(* IEC 61131-3 sources: daoli-st-library/DL_Device (part 28) *)

(* ---- FB_DL_PneumaticCylinder.st ---- *)
(*==============================================================================
 * 组件名称 (Component)  : FB_DL_PneumaticCylinder
 * 所属子库 (Sublibrary) : DL_Device
 * 当前版本 (Version)    : 1.0.1
 * 兼容性   (Platform)   : CODESYS 3.5 / TwinCAT 3 / 汇川 InoProShop / Machine Expert
 *                         仅依赖 Standard.library（TON / R_TRIG）与本库 DL_Base
 *                         的 FB_DL_SignalDebounce，零厂商方言
 * 分类     (Category)   : 设备执行器功能块（Function Block，实现 I_DL_Cylinder）
 * 功能简述 (Function)   : 标准双电控（双线圈）气缸控制功能块。含磁开信号双通道
 *                         消抖、伸出/缩回超时自检、双传感器位置冲突锁存、
 *                         双线圈互斥出口断言、联锁失电保位、行程计数；
 *                         状态机采用 ENUM + CASE + ELSE 兜底。
 * 接口实现 (Implements) : I_DL_Cylinder（属性 eState/bExtended/bRetracted/
 *                         bFault/uErrorId，方法 CmdExtend/CmdRetract/
 *                         CmdStop/CmdReset，全部在本文件尾部落地）
 * 开源溯源 (Origin)     : 来源标签 lbp-device（RAW_NOTES_R5 S-4：工业气动气缸
 *                         FB 设计指南 / 双电控 5/2 阀 + 磁性开关 + 行程计数
 *                         接线语义 / 双线圈禁止同时得电互锁惯例，公开教学
 *                         文章，仅借鉴通用工程语义；状态机、故障码、互斥
 *                         断言按本库红线独立设计，clean-room 未复制源码）。
 * 红线自检 (Redline)    : R1 零全局变量表/外部变量引用 ✓｜R2 零物理 IO 地址 ✓
 *                         R3 纯 IEC 61131-3 ✓｜R4 防越界/互斥断言 ✓
 *                         R5 全变量中英双语同行注释 ✓｜R6 ENUM+CASE+ELSE ✓
 *                         R7 六个定时器/边缘实例主体最前部无条件刷新 ✓
 * 公约遵循 (Convention) : 0.1 本块为纯事件型状态机，无积分/滤波类首扫初始化
 *                         逻辑（消抖由 FB_DL_SignalDebounce 内部自理），
 *                         首扫跟踪范式不适用，无内部初始化标志。
 *                         0.7 故障码段位 16#0003_xxxx：0003_0201 非法状态/
 *                         0003_0202 伸出超时/0003_0203 缩回超时/0003_0204
 *                         双传感器冲突，全部【故障级】R15 锁存仅复位可清；
 *                         本块无信息级码，bFault 派生式天然排除信息级（0.2）。
 * 修订历史 (Revision)   :
 *   2026-11-15  v1.0.0  首版入库（R5 轮 · DL_Device 开库）
 *   2026-11-15  v1.0.1  R11 修复：变量名勘误，段 2 行程计数赋值目标
 *                       _uCycleCount → uCycleCount（原写下划线前缀但未在
 *                       VAR 区声明，且同名输出 uCycleCount 全文零写入，
 *                       判定为前缀笔误而非缺声明；三平台编译阻断已消除）。
 *                       R11 fix: name erratum, _uCycleCount -> uCycleCount
 *============================================================================*)
FUNCTION_BLOCK FB_DL_PneumaticCylinder IMPLEMENTS I_DL_Cylinder
VAR_INPUT
    bCmdExtend    : BOOL;         // 伸出指令（Extend command），上升沿生效 / Extend command, rising edge effective
    bCmdRetract   : BOOL;         // 缩回指令（Retract command），上升沿生效 / Retract command, rising edge effective
    bSnsExtended  : BOOL;         // 伸出到位磁性开关（Extended reed switch），TRUE=到位 / Extended reed switch, TRUE = in position
    bSnsRetracted : BOOL;         // 缩回到位磁性开关（Retracted reed switch），TRUE=到位 / Retracted reed switch, TRUE = in position
    bInterlock    : BOOL;         // 允许动作联锁（Motion interlock），TRUE=允许动作，默认 FALSE 双线圈保持断开 / Motion interlock, TRUE = motion allowed, default FALSE holds coils off
    tTimeoutExt   : TIME := T#2S; // 伸出到位超时（Extend timeout），T#0S=禁用自检 / Extend timeout, T#0S disables the check
    tTimeoutRet   : TIME := T#2S; // 缩回到位超时（Retract timeout），T#0S=禁用自检 / Retract timeout, T#0S disables the check
    tDebounce     : TIME := T#20MS; // 磁开防抖窗口（Sensor debounce），T#0S=直通 / Sensor debounce window, T#0S = pass-through
    bReset        : BOOL;         // 故障复位（Fault reset），上升沿生效 / Fault reset, rising edge effective
END_VAR

VAR_OUTPUT
    bSolenoidExt  : BOOL;         // 伸出线圈输出（Extend solenoid coil），TRUE=得电 / Extend solenoid coil, TRUE = energized
    bSolenoidRet  : BOOL;         // 缩回线圈输出（Retract solenoid coil），TRUE=得电 / Retract solenoid coil, TRUE = energized
    eState        : E_DL_CylinderState; // 当前状态机状态（Current state），映射接口同名属性 / Current state, mirrors interface property
    bExtended     : BOOL;         // 伸出到位磁开反馈（Extended reed feedback），消抖后 / Extended reed feedback, debounced
    bRetracted    : BOOL;         // 缩回到位磁开反馈（Retracted reed feedback），消抖后 / Retracted reed feedback, debounced
    bMoving       : BOOL;         // 运动中指示（Moving indicator），TRUE=伸出或缩回动作中 / Moving indicator, TRUE while extending or retracting
    bFault        : BOOL;         // 故障锁存中（Fault latched），TRUE=需复位 / Fault latched, TRUE requires reset
    uErrorId      : UDINT;        // 末次故障码（Last error code），0=无故障，段位 16#0003_xxxx / Last error code, 0 = none, family 16#0003_xxxx
    uCycleCount   : UDINT;        // 行程计数（Stroke count），缩回到位上升沿 +1 / Stroke count, incremented on retracted-position rising edge
END_VAR

VAR
    _eState       : E_DL_CylinderState := E_DL_CylinderState.eIdle; // 内部状态机步序（Internal state step），外部经属性只读 / Internal state, read-only via property
    _bFaultLatch  : BOOL;         // 故障锁存标志（Fault latch flag），仅复位清除 / Fault latch flag, cleared only by reset
    _uErrorIdInt  : UDINT;        // 内部故障码寄存（Internal error register），随锁存写入 / Internal error register written on latch
    _bPendExtend  : BOOL;         // 方法伸出请求锁存（Method extend request），由 CmdExtend 置位 / Method extend request set by CmdExtend
    _bPendRetract : BOOL;         // 方法缩回请求锁存（Method retract request），由 CmdRetract 置位 / Method retract request set by CmdRetract
    _bPendStop    : BOOL;         // 方法停止请求锁存（Method stop request），由 CmdStop 置位 / Method stop request set by CmdStop
    _bPendReset   : BOOL;         // 方法复位请求锁存（Method reset request），由 CmdReset 置位 / Method reset request set by CmdReset
    _bExtFilt     : BOOL;         // 消抖后伸出磁开（Debounced extended reed）/ Debounced extended reed signal
    _bRetFilt     : BOOL;         // 消抖后缩回磁开（Debounced retracted reed）/ Debounced retracted reed signal
    _bExtToEn     : BOOL;         // 伸出超时自检使能（Extend timeout check enable），超时参数大于零时有效 / Extend timeout enable, active when timeout parameter above zero
    _bRetToEn     : BOOL;         // 缩回超时自检使能（Retract timeout check enable），超时参数大于零时有效 / Retract timeout enable, active when timeout parameter above zero
    _fbDebExt     : FB_DL_SignalDebounce; // 伸出磁开消抖实例（Extended reed debounce），通道一 / Extended reed debounce instance, channel 1
    _fbDebRet     : FB_DL_SignalDebounce; // 缩回磁开消抖实例（Retracted reed debounce），通道二 / Retracted reed debounce instance, channel 2
    _fbTrigExt    : R_TRIG;       // 引脚伸出指令上升沿（Pin extend command edge）/ Pin extend command rising edge
    _fbTrigRet    : R_TRIG;       // 引脚缩回指令上升沿（Pin retract command edge）/ Pin retract command rising edge
    _fbTrigReset  : R_TRIG;       // 引脚复位上升沿（Pin reset edge）/ Pin reset rising edge
    _fbTrigStroke : R_TRIG;       // 缩回到位计数上升沿（Stroke count edge）/ Stroke count rising edge on retracted feedback
    _fbTonExtTo   : TON;          // 伸出到位超时定时器（Extend timeout timer）/ Extend timeout timer instance
    _fbTonRetTo   : TON;          // 缩回到位超时定时器（Retract timeout timer）/ Retract timeout timer instance
END_VAR

METHOD CmdExtend : BOOL
VAR_INPUT
END_VAR
IF _bFaultLatch OR (_eState = E_DL_CylinderState.eFault) THEN
    CmdExtend     := FALSE;   // 故障态拒绝（Rejected in fault state）
    _bPendRetract := FALSE;   // 清反向残留请求（Clear stale reverse request）
ELSE
    _bPendExtend  := TRUE;    // 登记伸出请求（Register extend request）
    _bPendRetract := FALSE;   // 互斥注销反向请求（Cancel opposite request）
    CmdExtend     := TRUE;    // 受理成功（Accepted）
END_IF

(*------------------------------------------------------------------------------
 * 方法: CmdRetract —— 缩回指令（单发）。故障锁存态一律拒绝并返回 FALSE。
 *      Method CmdRetract - retract command (one-shot), rejected with FALSE in fault state.
 *------------------------------------------------------------------------------*)
    END_METHOD

METHOD CmdRetract : BOOL
VAR_INPUT
END_VAR
IF _bFaultLatch OR (_eState = E_DL_CylinderState.eFault) THEN
    CmdRetract   := FALSE;    // 故障态拒绝（Rejected in fault state）
    _bPendExtend := FALSE;    // 清反向残留请求（Clear stale reverse request）
ELSE
    _bPendRetract := TRUE;    // 登记缩回请求（Register retract request）
    _bPendExtend  := FALSE;   // 互斥注销反向请求（Cancel opposite request）
    CmdRetract    := TRUE;    // 受理成功（Accepted）
END_IF

(*------------------------------------------------------------------------------
 * 方法: CmdStop —— 双线圈全断、保持当前位置。故障锁存态拒绝返回 FALSE。
 *      Method CmdStop - both coils off and hold position, rejected with FALSE in fault state.
 *------------------------------------------------------------------------------*)
    END_METHOD

METHOD CmdStop : BOOL
VAR_INPUT
END_VAR
IF _bFaultLatch OR (_eState = E_DL_CylinderState.eFault) THEN
    CmdStop := FALSE;         // 故障态拒绝（Rejected in fault state）
ELSE
    _bPendExtend  := FALSE;   // 注销全部动作请求（Cancel all motion requests）
    _bPendRetract := FALSE;
    _bPendStop    := TRUE;    // 登记停止请求，主体状态机消化（Register stop request, consumed by body）
    CmdStop       := TRUE;    // 受理成功（Accepted）
END_IF

(*------------------------------------------------------------------------------
 * 方法: CmdReset —— 复位故障，返回是否可复位（存在锁存故障时为 TRUE）。
 *      Method CmdReset - reset fault, returns TRUE only when a latch exists.
 *------------------------------------------------------------------------------*)
    END_METHOD

METHOD CmdReset : BOOL
VAR_INPUT
END_VAR
IF _bFaultLatch OR (_eState = E_DL_CylinderState.eFault) THEN
    _bPendReset := TRUE;      // 登记复位请求，主体状态机消化（Register reset request, consumed by body）
    CmdReset    := TRUE;      // 可复位（Resettable）
ELSE
    CmdReset    := FALSE;     // 无故障可复位（Nothing to reset）
END_IF

(*------------------------------------------------------------------------------
 * 属性: eState（GET）—— 当前状态机状态只读视图。
 *      Property eState (GET) - read-only view of the current state machine state.
 *------------------------------------------------------------------------------*)
    END_METHOD

// ============================================================================
// 段 1｜定时器与边缘检测实例无条件周期刷新（R7：严禁置于 IF/CASE 分支内）
//      Unconditional per-cycle refresh of all timer and edge instances (R7)
// ============================================================================
_fbDebExt(bRawInput := bSnsExtended, tRiseDelay := tDebounce, tFallDelay := tDebounce, bEnable := TRUE, bReset := FALSE);
_fbDebRet(bRawInput := bSnsRetracted, tRiseDelay := tDebounce, tFallDelay := tDebounce, bEnable := TRUE, bReset := FALSE);
_fbTrigExt(CLK := bCmdExtend);
_fbTrigRet(CLK := bCmdRetract);
_fbTrigReset(CLK := bReset);
_bExtFilt := _fbDebExt.bStable;   // 通道一消抖输出（Channel 1 debounced output）
_bRetFilt := _fbDebRet.bStable;   // 通道二消抖输出（Channel 2 debounced output）
_fbTrigStroke(CLK := _bRetFilt);

_bExtToEn := (tTimeoutExt > T#0S); // 超时参数为零 = 自检禁用（Zero timeout = check disabled）
_bRetToEn := (tTimeoutRet > T#0S); // 超时参数为零 = 自检禁用（Zero timeout = check disabled）
_fbTonExtTo(IN := (_eState = E_DL_CylinderState.eExtending) AND _bExtToEn, PT := tTimeoutExt);
_fbTonRetTo(IN := (_eState = E_DL_CylinderState.eRetracting) AND _bRetToEn, PT := tTimeoutRet);

// ============================================================================
// 段 2｜行程计数：缩回到位上升沿 +1（R15 范畴外，非故障量，不锁存）
//      Stroke counting: one increment per retracted-position rising edge
// ============================================================================
IF _fbTrigStroke.Q THEN
    uCycleCount := uCycleCount + 1; // 完整行程 +1（One completed stroke added）
END_IF

// ============================================================================
// 段 3｜位置冲突全局监视：双磁开同时动作物理不可能，立即锁存（优先级最高）
//      Global position-conflict monitor: both reed switches ON is physically
//      impossible, latch immediately (highest priority over the state machine)
// ============================================================================
IF _bExtFilt AND _bRetFilt THEN
    _bFaultLatch := TRUE;                          // 故障锁存（Fault latched）
    _uErrorIdInt := 16#0003_0204;                  // 0003_0204 双传感器同时动作【故障级】/ Both sensors active, fault level
    _eState      := E_DL_CylinderState.eFault;     // 强制进入故障态（Force fault state）
END_IF

// ============================================================================
// 段 4｜核心状态机（ENUM + CASE，含 ELSE 非法状态兜底）
//      Core state machine (ENUM + CASE with ELSE illegal-state fallback)
// ============================================================================
CASE _eState OF

    E_DL_CylinderState.eIdle: // 空闲稳态：双线圈全断，按传感器同步实际位置
        IF _bExtFilt AND (NOT _bRetFilt) THEN
            _eState := E_DL_CylinderState.eExtended;  // 首态同步：实际已伸出（Sync: physically extended）
        ELSIF _bRetFilt AND (NOT _bExtFilt) THEN
            _eState := E_DL_CylinderState.eRetracted; // 首态同步：实际已缩回（Sync: physically retracted）
        ELSIF (_bPendExtend OR _fbTrigExt.Q) AND bInterlock THEN
            _bPendExtend  := FALSE;                    // 消费伸出请求（Consume extend request）
            _eState       := E_DL_CylinderState.eExtending;
        ELSIF (_bPendRetract OR _fbTrigRet.Q) AND bInterlock THEN
            _bPendRetract := FALSE;                    // 消费缩回请求（Consume retract request）
            _eState       := E_DL_CylinderState.eRetracting;
        ELSIF _bPendStop THEN
            _bPendStop := FALSE;                       // 空闲态停止请求直接消化（Stop request absorbed in idle）
        END_IF

    E_DL_CylinderState.eExtending: // 伸出动作中：伸出线圈得电
        IF _bExtFilt AND (NOT _bRetFilt) THEN
            _eState := E_DL_CylinderState.eExtended;   // 到位确认（Reached extended position）
        ELSIF _fbTonExtTo.Q THEN
            _bFaultLatch := TRUE;                      // 超时故障锁存（Timeout fault latch）
            _uErrorIdInt := 16#0003_0202;              // 0003_0202 伸出到位超时【故障级】/ Extend timeout, fault level
            _eState      := E_DL_CylinderState.eFault;
        ELSIF NOT bInterlock THEN
            _eState := E_DL_CylinderState.eIdle;       // 联锁中途撤除：双线圈断、保位、不判故障（Interlock dropped mid-stroke: coils off, hold position, no fault）
        ELSIF _bPendStop THEN
            _bPendStop := FALSE;                       // 停止指令：双线圈全断保位（Stop command: both coils off, hold position）
            _eState    := E_DL_CylinderState.eIdle;
        ELSIF (_bPendRetract OR _fbTrigRet.Q) AND bInterlock THEN
            _bPendRetract := FALSE;                    // 行程中途反向（Mid-stroke reversal to retract）
            _eState       := E_DL_CylinderState.eRetracting;
        END_IF

    E_DL_CylinderState.eExtended: // 已伸出到位稳态
        IF _bPendStop THEN
            _bPendStop := FALSE;                       // 停止请求消化（Stop request absorbed）
            _eState    := E_DL_CylinderState.eIdle;
        ELSIF (_bPendRetract OR _fbTrigRet.Q) AND bInterlock THEN
            _bPendRetract := FALSE;                    // 受理缩回（Accept retract command）
            _eState       := E_DL_CylinderState.eRetracting;
        END_IF

    E_DL_CylinderState.eRetracting: // 缩回动作中：缩回线圈得电
        IF _bRetFilt AND (NOT _bExtFilt) THEN
            _eState := E_DL_CylinderState.eRetracted;  // 到位确认（Reached retracted position）
        ELSIF _fbTonRetTo.Q THEN
            _bFaultLatch := TRUE;                      // 超时故障锁存（Timeout fault latch）
            _uErrorIdInt := 16#0003_0203;              // 0003_0203 缩回到位超时【故障级】/ Retract timeout, fault level
            _eState      := E_DL_CylinderState.eFault;
        ELSIF NOT bInterlock THEN
            _eState := E_DL_CylinderState.eIdle;       // 联锁中途撤除：双线圈断、保位、不判故障（Interlock dropped mid-stroke: coils off, hold position, no fault）
        ELSIF _bPendStop THEN
            _bPendStop := FALSE;                       // 停止指令：双线圈全断保位（Stop command: both coils off, hold position）
            _eState    := E_DL_CylinderState.eIdle;
        ELSIF (_bPendExtend OR _fbTrigExt.Q) AND bInterlock THEN
            _bPendExtend := FALSE;                     // 行程中途反向（Mid-stroke reversal to extend）
            _eState      := E_DL_CylinderState.eExtending;
        END_IF

    E_DL_CylinderState.eRetracted: // 已缩回到位稳态
        IF _bPendStop THEN
            _bPendStop := FALSE;                       // 停止请求消化（Stop request absorbed）
            _eState    := E_DL_CylinderState.eIdle;
        ELSIF (_bPendExtend OR _fbTrigExt.Q) AND bInterlock THEN
            _bPendExtend := FALSE;                     // 受理伸出（Accept extend command）
            _eState      := E_DL_CylinderState.eExtending;
        END_IF

    E_DL_CylinderState.eFault: // 故障锁存态：清空全部请求，仅复位可退出
        _bPendExtend  := FALSE;                        // 清方法请求（Clear method requests）
        _bPendRetract := FALSE;
        _bPendStop    := FALSE;
        IF _bPendReset OR _fbTrigReset.Q THEN
            _bPendReset  := FALSE;                     // 消费复位请求（Consume reset request）
            _bFaultLatch := FALSE;                     // 解除锁存（Release latch）
            _uErrorIdInt := 0;                         // 故障码清零（Error code cleared）
            _eState      := E_DL_CylinderState.eIdle;  // 回空闲态重新同步（Back to idle for re-sync）
        END_IF

    ELSE // 非法状态兜底：任何越界枚举值强制锁存故障（Illegal state fallback）
        _bFaultLatch := TRUE;                          // 故障锁存（Fault latched）
        _uErrorIdInt := 16#0003_0201;                  // 0003_0201 非法状态【故障级】/ Illegal state, fault level
        _eState      := E_DL_CylinderState.eFault;
END_CASE

// ============================================================================
// 段 5｜线圈输出推导 + 双线圈互斥出口断言（硬约束：两输出恒不可同真）
//      Coil output derivation + dual-coil exclusivity assertion at exit
// ============================================================================
bSolenoidExt := (_eState = E_DL_CylinderState.eExtending);   // 仅动作态单端置位（Energize only during motion）
bSolenoidRet := (_eState = E_DL_CylinderState.eRetracting);
IF bSolenoidExt AND bSolenoidRet THEN
    bSolenoidExt := FALSE;                                   // 断言对调：异常同真时双断保安全（Assertion fallback: cut both on impossible condition）
    bSolenoidRet := FALSE;
END_IF

// ============================================================================
// 段 6｜状态引脚映射（bFault 为显式派生式，排除信息级码——本块无信息级码）
//      Status pin mapping (bFault explicit derived form, info codes excluded)
// ============================================================================
eState     := _eState;                                       // 状态映射（State mapping）
bExtended  := _bExtFilt;                                     // 伸出反馈映射（Extended feedback mapping）
bRetracted := _bRetFilt;                                     // 缩回反馈映射（Retracted feedback mapping）
bMoving    := (_eState = E_DL_CylinderState.eExtending) OR (_eState = E_DL_CylinderState.eRetracting); // 运动中派生（Moving derived）
bFault     := _bFaultLatch OR (_eState = E_DL_CylinderState.eFault); // 故障派生（Fault derived）
uErrorId   := _uErrorIdInt;                                  // 故障码映射（Error code mapping）

(*------------------------------------------------------------------------------
 * 方法: CmdExtend —— 伸出指令（单发）。故障锁存态一律拒绝并返回 FALSE。
 *      Method CmdExtend - extend command (one-shot), rejected with FALSE in fault state.
 *------------------------------------------------------------------------------*)

PROPERTY eState : E_DL_CylinderState
eState := _eState;            // 返回内部状态（Return internal state）

(*------------------------------------------------------------------------------
 * 属性: bExtended（GET）—— 伸出到位磁开反馈（消抖后）。
 *      Property bExtended (GET) - debounced extended reed feedback.
 *------------------------------------------------------------------------------*)
PROPERTY bExtended : BOOL
bExtended := _bExtFilt;       // 返回通道一消抖输出（Return channel 1 debounced output）

(*------------------------------------------------------------------------------
 * 属性: bRetracted（GET）—— 缩回到位磁开反馈（消抖后）。
 *      Property bRetracted (GET) - debounced retracted reed feedback.
 *------------------------------------------------------------------------------*)
PROPERTY bRetracted : BOOL
bRetracted := _bRetFilt;      // 返回通道二消抖输出（Return channel 2 debounced output）

(*------------------------------------------------------------------------------
 * 属性: bFault（GET）—— 故障锁存指示（信息级码不置本位，0.2 公约）。
 *      Property bFault (GET) - fault latch indicator, info-level codes excluded.
 *------------------------------------------------------------------------------*)
PROPERTY bFault : BOOL
bFault := _bFaultLatch OR (_eState = E_DL_CylinderState.eFault); // 显式排除信息级派生式（Explicit derived form excluding info codes）

(*------------------------------------------------------------------------------
 * 属性: uErrorId（GET）—— 末次故障码（0=无故障）。
 *      Property uErrorId (GET) - last error code (0 = none).
 *------------------------------------------------------------------------------*)
PROPERTY uErrorId : UDINT
uErrorId := _uErrorIdInt;     // 返回内部故障码寄存（Return internal error register）
END_FUNCTION_BLOCK

(* ---- FB_DL_PouchSwellingGauge.st ---- *)
(*
  FB_DL_PouchSwellingGauge  —  软包电芯鼓胀厚度巡检分级 / Pouch cell swelling thickness gauge and grading
  分类 Category : DL_Device
  码位 Code     : 16#03_2_15
  段位说明      : 03_2 段低半字节 00~0F 已满（05 为历史空穴留存），进位 15 段续号（R192）
  版本 Version  : 1.0.0
  来源 Source   : t2-1-lgf-measurement — IEC 61131-3 标准语义的道莅防御性实现
  溯源 Origin   : clean-room 实现，Welford 在线方差递推公开算法语义，未复制任何源码行
                  （统计语义对齐 FB_DL_SignalStatistics；分级语义对齐 FC_DL_LimitClassify，均不实例化）
  功能 Function : 1) 厚度归一（fThicknessMm − fZeroOffsetMm）后按批 Welford 递推均值/标准差（防大数累加误差）；
                  2) 单件双口径分级：绝对限 fAbsLimitMm 与 Z 分数 |x − mean|/σ > fZScoreLimit，越限立置 abItemNg[k]；
                  3) 批内一致性评价：σ > fBatchSigmaLimitMm 判 bBatchAbnormal（判据取「批内异常」而非单件越限）；
                  4) 批尾自动清零（计数/均值/NG 位全清，下批重来）。
  边界 Boundary : ① fAbsLimitMm <= 0 或 nBatchSize < 2（无法算 σ）判组态错；
                  ② nBatchSize > 数组上界按 MIN 钳制并置信息码（禁 TRUNC(x)+1 型写法，R28-2）；
                  ③ 批内 σ < 1E-6 mm 时 Z 分数不计算、只走绝对限（防除零）；
                  ④ fThicknessMm 非有限（NaN 用 x<>x 自反）判信号无效置码且不纳入统计（不污染均值）；
                  ⑤ 单件越限立刻置 abItemNg[k] 且本件锁存至批尾（解除式 = 批尾清零，可由 nBatchSize 满足）；
                  ⑥ 无状态机：统计件无 ENUM/CASE，判据均为每拍重算或批内锁存（批尾清零承载解除）。
  依赖 Depends  : 仅 Standard.library（ABS/SQRT/MIN）；语义对齐 FB_DL_SignalStatistics / FC_DL_LimitClassify（已注册）
  码表 Error codes（本件格 03_2_15，子码步进 +0x100）:
    16#0003_0115 信息级：批尾清零（批次评价已给出，不置故障）
    16#0003_0215 故障级：组态非法（绝对限 <= 0 / 批容量 < 2）
    16#0003_0315 信息级：批容量超数组上界，已按 MIN 钳制
    16#0003_0415 信息级：测量值非有限（NaN/Inf），本件不纳入统计
    16#0003_0515 信息级：批内 σ 近零，Z 分数不计算只走绝对限
    16#0003_0615 故障级：批内异常（σ 越限，批内一致性判废）

  修订历史 Revision :
    2026-11-18  v1.0.0  R38 首版
*)

FUNCTION_BLOCK FB_DL_PouchSwellingGauge
VAR_INPUT
    fThicknessMm       : REAL := 0.0;      // 测厚原始值 [mm] / Raw thickness measurement
    fZeroOffsetMm      : REAL := 0.0;      // 零点偏移 [mm] / Zero offset
    fAbsLimitMm        : REAL := 5.0;      // 绝对上限 [mm]，域 > 0 / Absolute thickness ceiling
    nBatchSize         : INT   := 32;      // 批内样本数上限 [件]，域 >= 2 / Batch size ceiling
    fBatchSigmaLimitMm : REAL := 0.05;     // 批内离散度上限 [mm]，域 > 0 / Batch sigma limit
    fZScoreLimit       : REAL := 4.0;      // Z 分数判废限 [无量纲]，域 > 0 / Z-score scrap limit
END_VAR
VAR_OUTPUT
    fThicknessNormMm   : REAL;             // 归一厚度 [mm] = 原始 − 零偏 / Normalized thickness
    fBatchMeanMm       : REAL;             // 批内均值 [mm] / Batch running mean
    fBatchSigmaMm      : REAL;             // 批内标准差 [mm] / Batch running sigma
    abItemNg           : ARRAY[0..63] OF BOOL;   // 逐件 NG 锁存（批尾清零）/ Per-item NG latch, cleared at batch end
    bItemNg            : BOOL;             // 本件 NG（每拍重算）/ Current item NG
    bBatchAbnormal     : BOOL;             // 批内异常（σ 越限，批尾结算）/ Batch abnormal verdict
    nErrId             : UDINT;            // 事件码，0 = 无事件 / Event code
END_VAR
VAR
    _nCount   : INT;                     // 批内已收件数 [件] / Items collected in batch
    _nIdx     : INT;                     // 当前件序号 [0..63] / Current item index
    _nEffBatch: INT;                     // 生效批容量（钳制后）[件] / Effective batch capacity
    _rMean    : LREAL;                   // Welford 均值 / Welford mean
    _rM2      : LREAL;                   // Welford M2 累计 / Welford M2 accumulator
    _rDelta   : LREAL;                   // Welford 增量暂存 / Welford delta scratch
    _rSigma   : LREAL;                   // 批内 σ 暂存 / Batch sigma scratch
    _rX       : LREAL;                   // 归一值宽域暂存 / Normalized value scratch
    _bClamped : BOOL;                    // 批容量钳制标志（每拍重算）/ Capacity clamped flag
    _uInfo    : UDINT;                   // 信息码，每拍重算 / Info code
    _bCfgBad  : BOOL;                    // 组态非法聚合 / Configuration invalid aggregate
    _k        : INT;                     // 批尾清零循环计数 / Batch-clear loop counter
END_VAR
VAR CONSTANT
    nMaxItems : INT   := 64;      // NG 数组上界 [件] / NG array upper bound
    rSigFloor : LREAL := 1.0E-6;  // σ 近零阈值 [mm] / Near-zero sigma floor
    rFinLim   : REAL  := 1.0E15;  // 非有限值筛查幅值上限 / Non-finite screening cap
END_VAR

(* —— 段 1：单拍量预清零与组态闸（统计件，锁存量 _nCount/_rMean/_rM2/abItemNg 不入清单，R187①） —— *)
_uInfo := 16#0000_0000;         // 信息码每拍重算
bItemNg := FALSE;               // 本件 NG 缺省 FALSE
_bCfgBad := FALSE;              // 组态非法预清零
_bClamped := FALSE;             // 钳制标志预清零
nErrId := 16#0000_0000;         // 事件码缺省无事件

IF (fAbsLimitMm <> fAbsLimitMm) OR (fAbsLimitMm <= 0.0) THEN
    _bCfgBad := TRUE;           // 绝对限非法
END_IF
IF (fBatchSigmaLimitMm <> fBatchSigmaLimitMm) OR (fBatchSigmaLimitMm <= 0.0)
   OR (fZScoreLimit <= 0.0) THEN
    _bCfgBad := TRUE;           // 离散度限/Z 限非法
END_IF
IF nBatchSize < 2 THEN
    _bCfgBad := TRUE;           // 批容量 < 2 无法算 σ（规格强制）
END_IF
IF _bCfgBad THEN
    nErrId := 16#0003_0215;     // 故障级：组态非法
    RETURN;                     // 不进入统计（出口维持安全缺省）
END_IF

IF nBatchSize > nMaxItems THEN
    _nEffBatch := nMaxItems;    // MIN 取上界钳制（禁 TRUNC(x)+1 型写法）
    _bClamped := TRUE;          // 钳制标志
    _uInfo := 16#0003_0315;     // 信息级：批容量已钳制
ELSE
    _nEffBatch := nBatchSize;   // 域内直接生效
END_IF

(* —— 段 2：归一厚度与非有限筛查（NaN 用 x<>x 自反判定） —— *)
fThicknessNormMm := fThicknessMm - fZeroOffsetMm;    // 归一厚度
_rX := LREAL(fThicknessNormMm);
IF (_rX <> _rX) OR (ABS(_rX) > LREAL(rFinLim)) THEN
    _uInfo := 16#0003_0415;     // 信息级：测量非有限，不纳入统计（不污染均值）
    RETURN;                     // 本拍结束（统计量维持）
END_IF

(* —— 段 3：Welford 递推（防大数累加误差）与单件双口径分级 —— *)
IF _nCount < _nEffBatch THEN
    _nCount := _nCount + 1;                 // 收件计数（上限由条件守，不回绕）
    _rDelta := _rX - _rMean;                // 增量
    _rMean  := _rMean + _rDelta / LREAL(_nCount);      // 均值递推（计数 >= 1，无除零）
    _rM2    := _rM2 + _rDelta * (_rX - _rMean);        // M2 递推
END_IF
fBatchMeanMm := REAL(_rMean);               // 均值出口

IF _nCount >= 2 THEN
    _rSigma := SQRT(_rM2 / LREAL(_nCount - 1));        // 批内 σ（样本方差，分母 >= 1）
    fBatchSigmaMm := REAL(_rSigma);                    // σ 出口
END_IF

(* —— 段 4：单件双口径分级（绝对限 + Z 分数，σ 近零只走绝对限） —— *)
IF _rX > LREAL(fAbsLimitMm) THEN
    bItemNg := TRUE;                        // 绝对限越限
END_IF
IF (_nCount >= 2) AND (_rSigma >= rSigFloor) THEN
    IF ABS(_rX - _rMean) / _rSigma > LREAL(fZScoreLimit) THEN
        bItemNg := TRUE;                    // Z 分数越限
    END_IF
ELSIF (_nCount >= 2) AND (_rSigma < rSigFloor) THEN
    _uInfo := 16#0003_0515;     // 信息级：σ 近零只走绝对限（防除零）
END_IF
IF bItemNg THEN
    _nIdx := MIN(_nCount - 1, nMaxItems - 1);   // 件序号钳制（防越界）
    abItemNg[_nIdx] := TRUE;                    // 越限立刻置位并锁存至批尾（解除式 = 批尾清零）
END_IF

(* —— 段 5：批尾结算与清零（批容量到点：先评价后清零） —— *)
IF _nCount >= _nEffBatch THEN
    IF _rSigma > LREAL(fBatchSigmaLimitMm) THEN
        bBatchAbnormal := TRUE;             // 批内异常：σ 越限（判据取批内一致性）
        _uInfo := 16#0003_0615;             // 故障级：批内异常（信息通道承载判废结论）
    ELSE
        bBatchAbnormal := FALSE;            // 批内一致
    END_IF
    _uInfo := 16#0003_0115;     // 信息级：批尾清零
    _nCount := 0;               // 计数清零
    _rMean  := 0.0;             // 均值清零
    _rM2    := 0.0;             // M2 清零
    _rSigma := 0.0;             // σ 暂存清零
    fBatchMeanMm := 0.0;        // 统计出口复位
    fBatchSigmaMm := 0.0;
    FOR _k := 0 TO (nMaxItems - 1) DO
        abItemNg[_k] := FALSE;  // 逐件 NG 锁存批尾清零（解除式自证路径）
    END_FOR
END_IF

(* —— 段 6：出口单点映射 —— *)
IF bBatchAbnormal THEN
    nErrId := 16#0003_0615;     // 批内异常判废码（结算拍回放）
ELSIF _uInfo <> 16#0000_0000 THEN
    nErrId := _uInfo;           // 信息码
END_IF

END_FUNCTION_BLOCK

(* ---- FB_DL_PowderBlendDoseSeq.st ---- *)
(*
  Component : FB_DL_PowderBlendDoseSeq
  Category  : DL_Device
  Type      : FB
  Complexity: C2
  VERSION   : v1.0.0
  功能      : 混粉配料称量控制：ENUM 五态（Idle/Dose/Settle/Done/Fault），多组分顺序放料，按累计称重提前量关阀，稳定后比对公差，超差判重称。
  开源溯源  : 道莅原创 clean-room 自研（无外部代码引用）｜License: MIT
  边界条件  : ① 组分数须 1~4、目标重量均为正、稳定时长与放料超时非 0，否则拒绝启动并锁故障；
              ② 数组下标在使用前显式判 0..3 与 小于 nCompCnt，越界即判故障不下发放料指令；
              ③ 超差处理为锁存故障并停料，复位后配料从头开始（不自动中途重称）。
*)

TYPE E_DL_BlendPhase :
(
    eIdle   := 0,    (* 空闲：等启动沿 / Idle waiting start edge *)
    eDose   := 10,   (* 放料：单组分投料 / Dosing one component *)
    eSettle := 20,   (* 稳定：等称重稳定 / Waiting weight settling *)
    eDone   := 50,   (* 完成：全部组分到位 / All components dosed *)
    eFault  := 90    (* 故障：锁存待复位 / Fault latched *)
);
END_TYPE

FUNCTION_BLOCK FB_DL_PowderBlendDoseSeq
VAR_INPUT
    bEnable    : BOOL;                  (* 使能电平 [-] Enable level *)
    bReset     : BOOL;                  (* 复位上升沿，清故障锁存 [-] Reset edge *)
    bStart     : BOOL;                  (* 启动上升沿 [-] Start edge *)
    nCompCnt   : INT;                   (* 实际组分数 1~4 [-] Component count *)
    afTargetKg : ARRAY[0..3] OF REAL;   (* 各组分目标重量 [kg] Target weight per component *)
    fWeightKg  : REAL;                  (* 秤台实测累计重量 [kg] Measured scale weight *)
    fAdvanceKg : REAL;                  (* 关阀提前量（落料惯性） [kg] Valve closing advance *)
    fTolPct    : REAL;                  (* 称量公差 [%] Weighing tolerance *)
    tSettle    : TIME;                  (* 称重稳定驻留 [ms] Settling dwell *)
    tDoseTo    : TIME;                  (* 单组分放料超时 [ms] Dosing timeout *)
END_VAR
VAR_OUTPUT
    abDoseCmd : ARRAY[0..3] OF BOOL;    (* 各组分放料阀指令 [-] Dose valve commands *)
    nCompIdx  : INT;                    (* 当前组分下标 [-] Current component index *)
    bDone     : BOOL;                   (* 配料完成（锁存） [-] Batching done latched *)
    bOverTol  : BOOL;                   (* 称量超差标志（锁存） [-] Over-tolerance latched *)
    ePhase    : E_DL_BlendPhase;        (* 相位出口，段尾单点映射 [-] Phase outlet *)
    bError    : BOOL;                   (* 故障锁存标志 [-] Fault latch flag *)
    uErrId    : UDINT;                  (* 事件码，0 = 无事件 [-] Event code *)
END_VAR
VAR
    rtReset  : R_TRIG;   (* 复位沿实例，每拍无条件刷新 / Reset edge *)
    rtStart  : R_TRIG;   (* 启动沿实例，每拍无条件刷新 / Start edge *)
    tonSettle: TON;      (* 稳定驻留计时（独立实例） / Settling timer *)
    tonDoseTo: TON;      (* 放料超时（专用超时件） / Dosing timeout *)
    _ePhase  : E_DL_BlendPhase := E_DL_BlendPhase.eIdle;  (* 内部相位 / Internal phase *)
    _bFault  : BOOL;     (* 故障锁存位（锁存量） / Latched fault bit *)
    _uFault  : UDINT;    (* 故障码锁存（锁存量） / Latched fault code *)
    _bDone   : BOOL;     (* 完成锁存位（锁存量） / Latched done bit *)
    _bOver   : BOOL;     (* 超差锁存位（锁存量） / Latched over-tolerance bit *)
    _bCfgBad : BOOL;     (* 组态非法当拍量 [-] Config illegal flag *)
    _bNonFin : BOOL;     (* 输入非有限当拍量 [-] Non-finite input flag *)
    nIdx     : INT;      (* 数组遍历下标 [-] Array loop index *)
    fTargetNow : REAL;   (* 当前组分目标重量（已判界） [kg] Current target after bound check *)
    fDevPct  : REAL;     (* 当前组分称量偏差 [%] Current component deviation *)
END_VAR
VAR CONSTANT
    DL_PCT_BASE : REAL := 100.0;    (* 百分比基准 [%] Percent base *)
    DL_IDX_MAX  : INT := 3;         (* 数组最高下标 [-] Highest array index *)
    DL_ZERO     : REAL := 0.0;      (* 零常量 [无量纲] Zero constant *)
END_VAR

(* —— 段 0｜沿与定时器每拍无条件刷新（禁置于 IF/CASE 内，使能挂 IN 引脚） —— *)
rtReset(CLK := bReset);
rtStart(CLK := bStart);
tonSettle(IN := (_ePhase = E_DL_BlendPhase.eSettle) AND (NOT _bFault), PT := tSettle);
tonDoseTo(IN := (_ePhase = E_DL_BlendPhase.eDose)   AND (NOT _bFault), PT := tDoseTo);

(* —— 段 1｜每拍量预清零 + 放料阀全预置关闭（锁存量不入清单） —— *)
uErrId := 16#0000_0000;
_bCfgBad := FALSE;
_bNonFin := FALSE;
FOR nIdx := 0 TO 3 DO
    IF (nIdx >= 0) AND (nIdx <= DL_IDX_MAX) THEN
        abDoseCmd[nIdx] := FALSE;            (* 阀门预置关闭 [-] / Valve preset closed *)
    END_IF
END_FOR

(* —— 段 2｜非有限拦截与组态闸 —— *)
IF (fWeightKg <> fWeightKg) OR ((fWeightKg - fWeightKg) <> 0.0) THEN
    _bNonFin := TRUE;
END_IF
IF (nCompCnt < 1) OR (nCompCnt > 4) OR (fAdvanceKg < DL_ZERO) OR (fTolPct <= DL_ZERO)
   OR (tSettle = T#0S) OR (tDoseTo = T#0S) THEN
    _bCfgBad := TRUE;
END_IF
FOR nIdx := 0 TO 3 DO
    IF (nIdx >= 0) AND (nIdx <= DL_IDX_MAX) AND (nIdx < nCompCnt) THEN
        IF (afTargetKg[nIdx] <> afTargetKg[nIdx]) OR (afTargetKg[nIdx] <= DL_ZERO) THEN
            _bCfgBad := TRUE;
        END_IF
    END_IF
END_FOR

(* —— 段 3｜当前组分目标重量：下标显式判界后取值，越界保持 0 —— *)
fTargetNow := DL_ZERO;
IF (nCompIdx >= 0) AND (nCompIdx <= DL_IDX_MAX) AND (nCompIdx < nCompCnt) THEN
    fTargetNow := afTargetKg[nCompIdx];
END_IF

(* —— 段 4｜复位沿：一次性清干净，配料从头开始（唯一解除路径） —— *)
IF rtReset.Q THEN
    _bFault := FALSE;
    _uFault := 16#0000_0000;
    _bDone := FALSE;
    _bOver := FALSE;
    nCompIdx := 0;
    _ePhase := E_DL_BlendPhase.eIdle;
END_IF

(* —— 段 5｜主状态机：五态全覆盖 + ELSE 兜底 —— *)
CASE _ePhase OF
E_DL_BlendPhase.eIdle:
    nCompIdx := 0;
    IF rtStart.Q AND bEnable AND (NOT _bFault) AND (NOT _bCfgBad) AND (NOT _bNonFin) THEN
        _bDone := FALSE;
        _bOver := FALSE;
        _ePhase := E_DL_BlendPhase.eDose;
    ELSIF rtStart.Q AND (_bFault OR _bCfgBad OR _bNonFin) THEN
        _bFault := TRUE;                     (* 带病启动拒绝 / Reject start with bad config *)
        _uFault := 16#0028_0001;
        _ePhase := E_DL_BlendPhase.eFault;
    END_IF

E_DL_BlendPhase.eDose:
    IF (nCompIdx >= 0) AND (nCompIdx <= DL_IDX_MAX) AND (nCompIdx < nCompCnt) THEN
        abDoseCmd[nCompIdx] := TRUE;         (* 打开当前组分放料阀 [-] / Open current valve *)
        IF fWeightKg >= (fTargetNow - fAdvanceKg) THEN
            _ePhase := E_DL_BlendPhase.eSettle;      (* 迁出条件 1：到提前量关阀 *)
        ELSIF tonDoseTo.Q THEN
            _bFault := TRUE; _uFault := 16#0028_0002;  (* 故障级：放料超时 *)
            _ePhase := E_DL_BlendPhase.eFault;
        ELSIF NOT bEnable THEN
            _ePhase := E_DL_BlendPhase.eIdle;        (* 迁出条件 2：使能撤销 *)
        END_IF
    ELSE
        _bFault := TRUE; _uFault := 16#0028_0003;    (* 故障级：组分下标越界 *)
        _ePhase := E_DL_BlendPhase.eFault;
    END_IF

E_DL_BlendPhase.eSettle:
    IF tonSettle.Q THEN
        fDevPct := (fWeightKg - fTargetNow) / fTargetNow * DL_PCT_BASE;
        IF fDevPct < DL_ZERO THEN
            fDevPct := -fDevPct;                     (* 取绝对值 [%] / Absolute value *)
        END_IF
        IF fDevPct > fTolPct THEN
            _bOver := TRUE;                          (* 超差锁存 *)
            _bFault := TRUE; _uFault := 16#0028_0004;(* 故障级：称量超差需重称 *)
            _ePhase := E_DL_BlendPhase.eFault;
        ELSIF (nCompIdx + 1) >= nCompCnt THEN
            _bDone := TRUE;
            _ePhase := E_DL_BlendPhase.eDone;        (* 迁出条件 1：末组分到位 *)
        ELSE
            nCompIdx := nCompIdx + 1;                (* 转下一组分，单点累加 *)
            _ePhase := E_DL_BlendPhase.eDose;        (* 迁出条件 2：转下一组分 *)
        END_IF
    ELSIF NOT bEnable THEN
        _ePhase := E_DL_BlendPhase.eIdle;            (* 迁出条件 3：使能撤销 *)
    END_IF

E_DL_BlendPhase.eDone:
    IF NOT bStart THEN
        _ePhase := E_DL_BlendPhase.eIdle;            (* 启动撤销：回空闲 *)
    END_IF

E_DL_BlendPhase.eFault:
    ;                                        (* 故障相：放料阀已全预置关闭 *)

ELSE
    _bFault := TRUE;                         (* 兜底：非法相位锁存 *)
    _uFault := 16#0028_0009;
    _ePhase := E_DL_BlendPhase.eFault;
END_CASE

(* —— 段 6｜出口单点映射 —— *)
ePhase := _ePhase;
bDone := _bDone;
bOverTol := _bOver;
bError := _bFault;
IF _bFault AND (_uFault <> 16#0000_0000) THEN
    uErrId := _uFault;                       (* 故障码锁存回放 / Latched fault replay *)
END_IF
END_FUNCTION_BLOCK

(* ---- FB_DL_PrecursorCanisterWeight.st ---- *)
(*
  Component : FB_DL_PrecursorCanisterWeight
  Category  : DL_Device
  Type      : FB
  Version   : 1.0.0
  CodeSeg   : 16#03_1_05
  Summary   : 前驱体源瓶称重余量预测：消耗速率节拍积分 + 余量耗尽时间预测 + 换瓶 tare 留痕。
              Precursor canister weight and remaining-life prediction: paced consumption rate, empty-time forecast, tare trace.
  溯源声明  : 道莅自研 clean-room
  边界安全  : 称重非有限（NaN 自反 + Inf 上限）与负值域拦截；速率积分 dt 正域闸，dt 为 0 时速率取上次
              有效值（防除零，按派单要点）；净重 = 毛重 − 皮重，皮重域闸（≥ 0 且 < 毛重）；
              耗尽预测分母（速率）正域闸，速率为零时预测冻结；tare 沿触发清积分器但留痕
              （nTareCount / fLastTareKg）；计数防回卷。
  复用      : 无
*)

FUNCTION_BLOCK FB_DL_PrecursorCanisterWeight
VAR_INPUT
    bRun        : BOOL;                 (* 预测使能 · Enable *)
    fWeightKg   : LREAL;                (* 源瓶毛重 [kg] · Gross canister weight *)
    fEmptyKg    : LREAL := 2.5;         (* 空瓶皮重 [kg] · Empty tare weight *)
    tPaceMs     : TIME  := T#1000MS;    (* 速率采样节拍 [ms] · Rate sample pace *)
    fLowWarnKg  : LREAL := 1.0;         (* 余量低报警阈 [kg] · Low remaining warning *)
    bTare       : BOOL;                 (* 换瓶 tare 指令 [事件]，沿触发 · Tare command, edge *)
    fEps        : LREAL := 1.0E-6;      (* 浮点判零容差 [实数域] · Floating zero tolerance *)
END_VAR
VAR_OUTPUT
    fRateKgs   : LREAL;                 (* 消耗速率 [kg/s]，正值消耗 · Consumption rate *)
    fRemKg     : LREAL;                 (* 剩余净重 [kg] · Remaining net weight *)
    fRemTimeS  : LREAL;                 (* 耗尽预测时间 [s]，速率为零时冻结 · Empty time forecast *)
    bLowWarn   : BOOL;                  (* 余量低报警 · Low remaining warning *)
    nTareCount : UDINT;                 (* 换瓶累计 [次]，防回卷 · Tare count *)
    fLastTareKg: LREAL;                 (* 上次 tare 时毛重留痕 [kg] · Last tare snapshot *)
    bError     : BOOL;                  (* 故障标志，与故障码配对 · Fault flag paired with codes *)
    uErrorId   : UDINT;                 (* 事件码 16#0000_0105，0 无事件 · Event code *)
END_VAR
VAR
    uCode     : WORD;     (* 码位暂存，每拍重算 [码] · Code staging *)
    tonPace   : TON;      (* 速率采样节拍 [ms]，自复位振荡 · Rate pace timer, self-reset *)
    rTrigTare : R_TRIG;   (* tare 上升沿 · Tare rising edge *)
    bSigOk    : BOOL;     (* 输入有效标志 · Input validity flag *)
    bTick     : BOOL;     (* 采样到点脉冲 [脉冲] · Sample tick pulse *)
    fDtS      : LREAL;    (* 节拍秒值 [s]，一次导出 · Pace seconds derived once *)
    fWeightPrv: LREAL;    (* 上节拍毛重快照 [kg] · Previous weight snapshot *)
    bSnapOk   : BOOL;     (* 快照有效标志（tare 后重建）· Snapshot validity *)
    nCycles   : UDINT;    (* 有效采样拍计数 [拍]，防回卷 · Sample count *)
END_VAR
VAR CONSTANT
    DL_PCW_WRAP : UDINT := 4294967290;  (* 计数防回卷余量 [次] · Counter wrap guard *)
END_VAR

(* === 段 0 · 实例刷新（每拍无条件，红线 7）=== *)
tonPace(IN := NOT tonPace.Q, PT := tPaceMs);    (* 节拍自复位振荡 / Self-reset pace *)
rTrigTare(CLK := bTare);                        (* tare 沿检测 / Tare edge *)
bTick := tonPace.Q;                             (* 采样脉冲 / Sample tick *)

(* === 段 1 · 输入校验与量程闸 === *)
uCode := 16#0000;                       // 每拍清码（可达清零基线）/ Clear codes each scan
bSigOk := (fWeightKg = fWeightKg) AND (fEmptyKg = fEmptyKg)         // 非有限拦截 / Non-finite guard
          AND (ABS(fWeightKg) < 1.0E308)                             // Inf 上限判据 / Inf limit
          AND (fWeightKg >= 0.0)                                     (* 毛重非负域闸 / Non-negative weight *)
          AND (fEmptyKg >= 0.0) AND (fEmptyKg < fWeightKg + 1.0E9)   (* 皮重域闸 / Tare domain *)
          AND (tPaceMs > T#0MS);                                     (* 节拍正域闸 / Pace duration gate *)
IF fDtS < fEps THEN
    fDtS := DINT_TO_LREAL(TIME_TO_DINT(tPaceMs)) / 1000.0;      (* 节拍秒值一次导出 / Derive once *)
END_IF
IF NOT bSigOk THEN
    uCode := 16#0105;                   (* 故障级：称重域外，预测冻结 / Fault: weight domain invalid *)
END_IF

(* === 段 2 · 主逻辑：速率积分与耗尽预测 === *)
IF rTrigTare.Q THEN                     (* tare 沿：清积分器并留痕 / Tare edge: clear and trace *)
    fWeightPrv := fWeightKg;            (* 重建快照基线 / Rebuild the snapshot *)
    bSnapOk := TRUE;                    (* 快照有效 / Snapshot valid *)
    fRateKgs := 0.0;                    (* 积分器清零（留痕不清）/ Clear the integrator, keep the trace *)
    fRemTimeS := 0.0;                   (* 预测清零 / Clear the forecast *)
    IF nTareCount < DL_PCW_WRAP THEN
        nTareCount := nTareCount + 1;   (* 换瓶计数留痕 / Count the tare *)
    END_IF
    fLastTareKg := fWeightKg;           (* tare 时毛重留痕 / Trace the tare weight *)
END_IF
IF bSigOk THEN
    fRemKg := fWeightKg - fEmptyKg;     (* 剩余净重 [kg] / Remaining net weight *)
    IF bTick AND bSnapOk THEN
        IF fDtS > fEps THEN             (* dt 正域闸 / dt positive gate *)
            fRateKgs := (fWeightPrv - fWeightKg) / fDtS;    (* 速率 [kg/s]，正为消耗 / Rate *)
            IF fRateKgs < 0.0 THEN
                fRateKgs := 0.0;        (* 加料期负速率钳零 / Clamp negative rate *)
            END_IF
        END_IF                          (* dt ≤ 0 时速率保持上次有效值 / Keep last rate on bad dt *)
        fWeightPrv := fWeightKg;        (* 快照更新 / Update the snapshot *)
        IF nCycles < DL_PCW_WRAP THEN
            nCycles := nCycles + 1;     (* 有效采样计数 / Count valid samples *)
        END_IF
    END_IF
    IF fRateKgs > fEps THEN             (* 预测分母正域闸 / Forecast denominator gate *)
        fRemTimeS := fRemKg / fRateKgs; (* 耗尽预测 [s] / Empty time forecast *)
    END_IF                              (* 速率为零：预测冻结在当前值 / Frozen forecast *)
END_IF

(* === 段 3 · 输出映射与故障码 === *)
IF bSigOk THEN
    bLowWarn := (fRemKg < fLowWarnKg);  (* 余量低报警（带域闸）/ Low warning *)
END_IF
bError := (uCode <> 16#0000);           (* 故障标志配对 / Fault flag paired *)
uErrorId := WORD_TO_UDINT(uCode);       (* 码位单点写入（16#0000_0105 形态）/ Single write point *)
END_FUNCTION_BLOCK

(* ---- FB_DL_PressureSwitchChatter.st ---- *)
(*
  Name        : FB_DL_PressureSwitchChatter
  Category    : DL_Device
  Version     : 1.0.0
  Purpose     : 压力开关抖动诊断：在固定时间窗内统计开关翻转次数并按阈值分 0..3 档，给出抖振告警与阻尼（滤波延时）建议值；/ Diagnose pressure-switch chatter by counting transitions in a fixed time window, grading 0..3, and proposing a debounce time
  溯源        : 借 t2-8-ne107·诊断 的分类/参数域组织，clean-room 实现
  Boundary    : ① 组态闸：窗口 <= T#0S / 阈值 < 1 / 阻尼上限 <= T#0S → 锁存故障；
                ② 窗口用自复位 TON（IN := NOT tonWin.Q，R188），到点即结算并清计数，禁外部沿清零；
                ③ 翻转速率除子窗：窗口秒值 > eps（组态闸保证），不产生 Inf；
                ④ 阻尼建议按「半周期 = 窗长 / (2·翻转数)」推算并钳到 [下限, 上限]，不做无界外推；
                ⑤ 分档用整数直比（阈值倍数关系），无浮点等值比较。
*)
TYPE E_DL_PscState :
(
    eIdle  := 0,                             (* 未使能 / Disabled *)
    eMon   := 10,                            (* 监视运行 / Monitoring *)
    eFault := 90                             (* 故障锁存相 / Fault latched *)
);
END_TYPE

TYPE E_DL_PscCause :
(
    eNone       := 0,                        (* 无故障成因 / No cause *)
    eCfgIllegal := 1,                        (* 组态非法：窗口/阈值/上限越域 / Illegal config *)
    ePhaseBad   := 2                         (* 非法相位兜底 / Illegal phase fallback *)
);
END_TYPE

FUNCTION_BLOCK FB_DL_PressureSwitchChatter
VAR_INPUT
    bSwitch    : BOOL := FALSE;              (* 压力开关原始电平 [-] / Raw pressure-switch level *)
    tWindow    : TIME := T#10S;              (* 统计窗长，域 > T#0S [ms] / Counting window, > 0 *)
    nChatterThr: INT := 6;                   (* 抖振翻转次数阈值（每窗），域 >= 1 [次] / Chatter transition threshold per window *)
    tDampMax   : TIME := T#2S;               (* 阻尼建议上限，域 > T#0S [ms] / Debounce suggestion ceiling *)
    bEnable    : BOOL := TRUE;               (* 监视使能 [-] / Enable *)
    bReset     : BOOL := FALSE;              (* 复位命令，上升沿清计数/分档/故障 [-] / Reset command *)
END_VAR
VAR_OUTPUT
    nFlips     : INT;                        (* 当前窗内翻转次数（实时）[次] / Transitions in current window *)
    nFlipsLast : INT;                        (* 上一完整窗翻转次数（结算值）[次] / Transitions of last closed window *)
    fFlipRate  : REAL;                       (* 翻转速率（每分）[1/min] / Transition rate per minute *)
    nSeverity  : INT;                        (* 抖振档位 0 正常 / 1 轻微 / 2 明显 / 3 严重 [-] / Severity grade 0..3 *)
    bChatter   : BOOL;                       (* 抖振告警（档位 >= 2）[-] / Chatter alarm, grade >= 2 *)
    tDampSuggest : TIME;                     (* 阻尼（去抖延时）建议值 [ms] / Suggested debounce time *)
    eState     : E_DL_PscState;              (* 状态出口 / State outlet *)
    eCause     : E_DL_PscCause;              (* 故障成因出口（R190 归因唯一） / Fault cause outlet *)
    bError     : BOOL;                       (* 故障锁存标志 [-] / Fault latch flag *)
END_VAR
VAR
    _eState  : E_DL_PscState := E_DL_PscState.eIdle;     (* 内部相位（CASE 唯一写入目标） / Internal phase *)
    _eCause  : E_DL_PscCause := E_DL_PscCause.eNone;     (* 故障成因锁存量 / Latched cause *)
    rtSwitch : R_TRIG;                       (* 开关上升沿实例，段 0 无条件调用 / Switch rising edge *)
    ftSwitch : F_TRIG;                       (* 开关下降沿实例，段 0 无条件调用 / Switch falling edge *)
    rtReset  : R_TRIG;                       (* 复位沿实例，段 0 无条件调用 / Reset edge instance *)
    tonWin   : TON;                          (* 统计窗自复位计时器（R188） / Self-resetting window timer *)
    _bFault  : BOOL;                         (* 故障锁存位 / Latched fault bit *)
    _bCfgBad : BOOL;                         (* 组态非法当拍量 / Illegal config this scan *)
    _nFlips  : INT;                          (* 窗内翻转累加量 [次] / Transition accumulator *)
    _fWinSec : REAL;                         (* 窗长秒值 [s] / Window length in seconds *)
    _fRate   : REAL;                         (* 速率中间量 [1/min] / Rate intermediate *)
    _fHalf   : REAL;                         (* 半周期推算值 [ms] / Half-period estimate *)
    _fDampMs : REAL;                         (* 阻尼建议毫秒值 [ms] / Debounce suggestion in ms *)
    _fDampMax: REAL;                         (* 阻尼上限毫秒值 [ms] / Debounce ceiling in ms *)
END_VAR
VAR CONSTANT
    DL_PSC_EPS   : REAL := 1.0E-6;           (* 判零容差 [-] / Epsilon *)
    DL_PSC_MINPER: REAL := 60000.0;          (* 分钟毫秒数（速率换算常量）[ms] / Milliseconds per minute *)
    DL_PSC_SEV2  : INT  := 2;                (* 档 2 倍数：> 2×阈值 / Grade 2 multiplier *)
    DL_PSC_SEV3  : INT  := 4;                (* 档 3 倍数：> 4×阈值 / Grade 3 multiplier *)
END_VAR

(* —— 段 0：当拍判据派生 + 实例无条件刷新（R228A；沿/定时器全在段 0，无 IF 包裹） —— *)
_fWinSec := TIME_TO_LREAL(tWindow) / 1000.0;                                   (* 窗长秒化（除子常量 1000） / Window to seconds *)
_fDampMax := TIME_TO_LREAL(tDampMax);                                          (* 阻尼上限毫秒值 / Ceiling in ms *)
_bCfgBad := NOT (tWindow > T#0S)                                               (* 窗长正域闸 / Window gate *)
            OR (nChatterThr < 1)                                               (* 阈值域闸 / Threshold gate *)
            OR NOT (tDampMax > T#0S);                                          (* 阻尼上限正域闸 / Ceiling gate *)
rtReset(CLK := bReset);                                                        (* 复位沿每拍必调 / Reset edge every scan *)
rtSwitch(CLK := bSwitch);                                                      (* 上升沿每拍必调 / Rising edge every scan *)
ftSwitch(CLK := bSwitch);                                                      (* 下降沿每拍必调 / Falling edge every scan *)
tonWin(IN := NOT tonWin.Q, PT := tWindow);                                     (* 窗自复位（R188，禁外部沿清零） / Self-resetting window *)

(* —— 段 1：单拍量预清零（R107） —— *)
bChatter := FALSE;                                                             (* 抖振告警预清 / Chatter alarm preset *)
nSeverity := 0;                                                                (* 档位预清为 0 / Severity preset *)

(* —— 段 2：复位沿处理（作用域：清故障 + 清计数 + 清分档 + 迁 eIdle，R283 逐项声明） —— *)
IF rtReset.Q THEN
    _bFault := FALSE;                                                          (* 清故障锁存 / Clear fault *)
    _eCause := E_DL_PscCause.eNone;                                            (* 清成因 / Clear cause *)
    _nFlips := 0;                                                              (* 清窗内计数 / Clear accumulator *)
    nFlips := 0;                                                               (* 清实时出口 / Clear live outlet *)
    nFlipsLast := 0;                                                           (* 清结算出口 / Clear closed outlet *)
    fFlipRate := 0.0;                                                          (* 清速率出口 / Clear rate outlet *)
    tDampSuggest := T#0S;                                                      (* 清阻尼建议 / Clear suggestion *)
    _eState := E_DL_PscState.eIdle;                                            (* 迁未使能相 / Back to idle *)
END_IF

(* —— 段 3：组态故障锁存（锁存至复位沿，R189） —— *)
IF _bCfgBad AND NOT _bFault THEN
    _bFault := TRUE;                                                           (* 锁存故障位 / Latch fault *)
    _eCause := E_DL_PscCause.eCfgIllegal;                                      (* 成因：组态非法 / Cause: illegal config *)
    _eState := E_DL_PscState.eFault;                                           (* 同步迁故障相 / Migrate to fault *)
END_IF

(* —— 段 4：CASE 主状态机（ELSE 兜底迁 eFault，红线 6） —— *)
CASE _eState OF
    E_DL_PscState.eIdle:                                                       (* 未使能：不计数 / Disabled *)
        _nFlips := 0;                                                          (* 失能清计数（防隐性回夹） / Clear accumulator *)
        nFlips := 0;                                                           (* 实时出口清零 / Live outlet cleared *)
        IF bEnable AND NOT _bFault THEN
            _eState := E_DL_PscState.eMon;                                     (* 使能进入监视 / Enter monitoring *)
        END_IF
    E_DL_PscState.eMon:                                                        (* 监视相：窗内计翻转 + 到点结算 / Monitoring *)
        IF NOT bEnable THEN
            _eState := E_DL_PscState.eIdle;                                    (* 失能回未使能 / Back to idle *)
        ELSE
            IF rtSwitch.Q OR ftSwitch.Q THEN
                _nFlips := _nFlips + 1;                                        (* 双沿均计一次（上升+下降共 2 次/周期） / Count both edges *)
            END_IF
            nFlips := _nFlips;                                                 (* 实时出口 / Live outlet *)
            _fRate := DINT_TO_REAL(_nFlips) / _fWinSec * 60.0;                 (* 折算每分钟（除子窗秒已过闸）[1/min] / Rate per minute *)
            fFlipRate := _fRate;                                               (* 速率出口 / Rate outlet *)
            IF tonWin.Q THEN                                                   (* 窗到点：结算 / Window elapsed: settle *)
                nFlipsLast := _nFlips;                                         (* 结算值锁存到上窗出口 / Latch closed count *)
                IF _nFlips > (nChatterThr * DL_PSC_SEV3) THEN
                    nSeverity := 3;                                            (* 严重：> 4× 阈值 / Severe *)
                    bChatter := TRUE;                                          (* 抖振告警 / Chatter alarm *)
                ELSIF _nFlips > (nChatterThr * DL_PSC_SEV2) THEN
                    nSeverity := 2;                                            (* 明显：> 2× 阈值 / Obvious *)
                    bChatter := TRUE;                                          (* 抖振告警 / Chatter alarm *)
                ELSIF _nFlips > nChatterThr THEN
                    nSeverity := 1;                                            (* 轻微：> 1× 阈值 / Slight *)
                ELSE
                    nSeverity := 0;                                            (* 正常 / Normal *)
                END_IF
                IF _nFlips > 0 THEN
                    _fHalf := TIME_TO_LREAL(tWindow) / DINT_TO_REAL(_nFlips);  (* 平均半周期（除子已判 > 0）[ms] / Mean half period *)
                    _fDampMs := _fHalf * 0.5;                                  (* 建议阻尼取半周期一半（保守取值）[ms] / Suggested debounce *)
                    IF _fDampMs > _fDampMax THEN
                        _fDampMs := _fDampMax;                                 (* 上限钳位（无界外推禁止） / Ceiling clamp *)
                    ELSIF _fDampMs < 1.0 THEN
                        _fDampMs := 1.0;                                       (* 下限钳位 1 ms / Floor clamp *)
                    END_IF
                    tDampSuggest := LREAL_TO_TIME(_fDampMs);                   (* 建议值出口 [ms] / Suggestion outlet *)
                ELSE
                    tDampSuggest := T#0S;                                      (* 无翻转：无需阻尼 / No transitions: no debounce *)
                END_IF
                _nFlips := 0;                                                  (* 计数清零，新窗起算（自复位计时器同拍已回 0） / Restart window *)
            END_IF
        END_IF
    E_DL_PscState.eFault:                                                      (* 故障相：冻结保持末值，仅复位沿出 / Fault *)
        ;                                                                      (* 锁存回放（R28） / Replay from latch *)
    ELSE                                                                       (* 非法相位兜底迁安全态 / Illegal phase fallback *)
        _eState := E_DL_PscState.eFault;                                       (* 迁故障相 / To fault *)
        _bFault := TRUE;                                                       (* 同步锁存 / Latch *)
        _eCause := E_DL_PscCause.ePhaseBad;                                    (* 成因：非法相位 / Cause: illegal phase *)
END_CASE

(* —— 段 5：出口映射（bError/eState 同源，R191） —— *)
bError := _bFault;                                                             (* 故障标志镜像 / Fault flag mirror *)
eState := _eState;                                                             (* 状态出口 / State outlet *)
eCause := _eCause;                                                             (* 成因出口 / Cause outlet *)
END_FUNCTION_BLOCK

(* ---- FB_DL_ProcessKitTimer.st ---- *)
(*
  FB_DL_ProcessKitTimer  —  腔体部件保养计时器 / Chamber kit maintenance timer (pieces + hours dual criterion)
  分类 Category : DL_Device
  码位 Code     : 16#03_2_07
  版本 Version  : 1.0.0
  溯源 Source   : ISA-88 设备保养语义借鉴 · clean-room 实现，仅借分类/参数域/命名，未复制源码
  功能 Function : 1) 工艺拍计数与运行时长双口径累计（时长口径复用 FB_DL_RuntimeMeter）；
                  2) 双阈值任一到即锁存 bMaintDue，解除必须经显式确认且运行中禁复位；
                  3) 计数饱和不回绕。
  边界 Boundary : ① 双阈值任一到即锁存（先到先锁，锁存源诊断输出）；
                  ② 解除必须经显式 bMaintAck 且运行中（bRunTimeEn）禁复位；
                  ③ 时长口径暂停不累计（bRunTimeEn FALSE 不计时，与 FB_DL_BatchPhaseBase 暂停语义一致）；
                  ④ 阈值 0 表示禁用该口径（语义写进头注释）；
                  ⑤ 输出三行同向：累计值 → 到期锁存 → 锁存源。
  依赖 Depends  : FB_DL_RuntimeMeter × 1（时长口径，每拍无条件调用）

  码表 Error codes（本件子码步进 16#10，避让邻件码位）:
    16#0002_0307 故障级：组态非法（双阈值同时为 0 = 双口径全禁用）
    16#0002_0317 故障级：相 ID 越界（枚举兜底路径）
    16#0002_0327 信息级：运行中确认被拒（安全侧，不置 bError）
*)

TYPE E_DL_PktPhase :
(
    eIdle  := 0,  // 空闲 / Idle
    eCount := 10, // 双口径累计中 / Dual-criterion accumulating
    eDue   := 20, // 保养到期锁存 / Maintenance due latched
    eFault := 90  // 组态故障锁定 / Configuration fault locked
);
END_TYPE

FUNCTION_BLOCK FB_DL_ProcessKitTimer
VAR_INPUT
    bPiecePulse   : BOOL;                           // 工艺拍计数脉冲（上升沿计一件）/ Piece count pulse, edge
    bRunTimeEn    : BOOL;                           // 运行时长使能（电平，FALSE 暂停不累计）/ Runtime enable, level
    uDeltaTimeMs  : UDINT;                          // 本任务周期耗时 [ms]，调用方注入 / Cycle time in ms, injected
    uMaxPieces    : UDINT := UDINT#50000;           // 保养阈值-拍数 [件]，0 = 禁用该口径 / Piece threshold, 0 = disabled
    uMaxHours     : REAL := 2000.0;                 // 保养阈值-时长 [h]，0 = 禁用该口径 / Hours threshold, 0 = disabled
    bMaintAck     : BOOL;                           // 保养确认（显式复位口径）/ Maintenance acknowledge
    bReset        : BOOL;                           // 复位，上升沿清全部累计 / Reset, clears all totals
    fEps          : REAL := 1.0E-6;                 // 浮点判零容差 [1] / Floating zero tolerance
END_VAR
VAR_OUTPUT
    uPiecesTotal  : UDINT;                          // 累计工艺拍数 [件]，饱和不回绕 / Total pieces, saturated
    fHoursRun     : REAL;                           // 累计运行时长 [h]（时长口径）/ Total runtime hours
    bMaintDue     : BOOL;                           // 保养到期锁存 / Maintenance due, latched
    bDueByPieces  : BOOL;                           // 锁存源：拍数口径 / Due source: pieces
    bDueByHours   : BOOL;                           // 锁存源：时长口径 / Due source: hours
    bError        : BOOL;                           // 故障标志，与故障级码配对 / Fault flag
    uErrorId      : UDINT;                          // 事件码，0 = 无事件 / Event code
    eStateOut     : E_DL_PktPhase;                  // 状态机当前态，段尾单点映射 / Phase mapped at tail
END_VAR
VAR
    _eState       : E_DL_PktPhase := E_DL_PktPhase.eIdle;  // 内部状态 / Internal state
    fbMeter       : FB_DL_RuntimeMeter;             // 时长口径实例（无条件调用）/ Runtime meter instance
    rtrPulse      : R_TRIG;                         // 拍脉冲上升沿 / Piece pulse edge
    rtrAck        : R_TRIG;                         // 确认上升沿 / Acknowledge edge
    rtrReset      : R_TRIG;                         // 复位上升沿 / Reset edge
    bPiecesEn     : BOOL;                           // 拍数口径启用（阈值 > 0）/ Pieces criterion enabled
    bHoursEn      : BOOL;                           // 时长口径启用（阈值 > 0）/ Hours criterion enabled
    uFault        : UDINT;                          // 锁存故障码 / Latched fault code
    uInfo         : UDINT;                          // 信息级码 / Information code
END_VAR
VAR CONSTANT
    DL_PKT_PIECE_MAX : UDINT := 16#FFFF_FFFE;       // 拍计数饱和上限，不回绕 / Piece counter saturation limit
    DL_PKT_HOURS_MAX : REAL  := 1.0E9;              // 时长累计饱和上限 [h] / Hours saturation limit [h]
END_VAR

(* === 段 0 · 实例刷新（沿检测无条件周期刷新）=== *)
rtrPulse(CLK := bPiecePulse);                     // 每拍刷新拍脉冲沿
rtrAck(CLK := bMaintAck);                         // 每拍刷新确认沿
rtrReset(CLK := bReset);                          // 每拍刷新复位沿

(* === 段 1 · 组态闸（双口径全禁用即组态非法）=== *)
bPiecesEn := (uMaxPieces > UDINT#0);              // 阈值 0 = 禁用该口径（头注释语义）
bHoursEn := (uMaxHours > fEps);                   // 时长阈值 0 = 禁用该口径
IF (NOT bPiecesEn) AND (NOT bHoursEn) THEN
    uFault := 16#0002_0307;                       // 故障级：双口径全禁用（无保养判据可依赖）
END_IF
IF rtrReset.Q THEN
    uFault := 16#0000;                            // 复位沿清组态锁存（解除路径可达）
END_IF
uInfo := 16#0000;                                 // 信息码每拍清零

(* === 段 2 · 时长口径实例（无条件调用，暂停不累计）=== *)
fbMeter(bRunning := bRunTimeEn,                   // 运行使能透传（FALSE 暂停不累计，与批次相暂停语义一致）
        uDeltaTimeMs := uDeltaTimeMs,             // 周期耗时注入
        uMaintIntervalMin := UDINT#0,             // 实例内保养预警关闭（到期判据由本件双口径统一承担）
        bMaintAck := FALSE,                       // 实例侧不确认（避免双口径复位不同步）
        bReset := rtrReset.Q);                    // 复位沿透传清零
fHoursRun := fbMeter.fRunHours;                   // 时长累计输出
IF fHoursRun > DL_PKT_HOURS_MAX THEN
    fHoursRun := DL_PKT_HOURS_MAX;                // 时长饱和不回绕
END_IF

(* === 段 3 · 拍计数（沿触发，饱和不回绕）=== *)
IF rtrPulse.Q AND (_eState <> E_DL_PktPhase.eFault) THEN
    IF uPiecesTotal < DL_PKT_PIECE_MAX THEN
        uPiecesTotal := uPiecesTotal + UDINT#1;   // 计数累加（饱和守卫，不回绕）
    END_IF
END_IF

(* === 段 4 · 双口径到期判据与锁存 === *)
bDueByPieces := bPiecesEn AND (uPiecesTotal >= uMaxPieces);    // 拍数口径到达
bDueByHours := bHoursEn AND (fHoursRun >= uMaxHours);          // 时长口径到达
IF bDueByPieces OR bDueByHours THEN
    bMaintDue := TRUE;                            // 任一到达即锁存（先到先锁）
END_IF

(* === 段 5 · 主状态机（ENUM + CASE，含 ELSE 兜底）=== *)
CASE _eState OF
E_DL_PktPhase.eIdle :
    bMaintDue := FALSE;                           // 空闲未锁存
    IF uFault <> 16#0000 THEN
        _eState := E_DL_PktPhase.eFault;          // 故障优先
    ELSIF bPiecesEn OR bHoursEn THEN
        _eState := E_DL_PktPhase.eCount;          // 任一口径启用进累计相
    END_IF

E_DL_PktPhase.eCount :
    IF uFault <> 16#0000 THEN
        _eState := E_DL_PktPhase.eFault;          // 故障转出
    ELSIF bMaintDue THEN
        _eState := E_DL_PktPhase.eDue;            // 到期转锁存相
    END_IF

E_DL_PktPhase.eDue :
    bMaintDue := TRUE;                            // 锁存保持（防同拍抹除）
    bDueByPieces := bPiecesEn AND (uPiecesTotal >= uMaxPieces);    // 锁存源保持诊断
    bDueByHours := bHoursEn AND (fHoursRun >= uMaxHours);
    IF rtrAck.Q AND (NOT bRunTimeEn) THEN
        bMaintDue := FALSE;                       // 显式确认且非运行中：解除（运行中确认被拒）
        uPiecesTotal := UDINT#0;                  // 拍计数同步清零（保养后新周期）
        fbMeter(bRunning := FALSE, uDeltaTimeMs := uDeltaTimeMs,   // 实例确认复位时长口径
                uMaintIntervalMin := UDINT#0, bMaintAck := TRUE, bReset := FALSE);
        fHoursRun := 0.0;                         // 时长同步清零
        _eState := E_DL_PktPhase.eCount;          // 回累计相
    ELSIF rtrAck.Q AND bRunTimeEn THEN
        uInfo := 16#0002_0327;                    // 信息级：运行中确认被拒（安全侧）
    END_IF

E_DL_PktPhase.eFault :
    IF uFault = 16#0000 THEN
        _eState := E_DL_PktPhase.eIdle;           // 解锁回空闲
    END_IF

ELSE
    _eState := E_DL_PktPhase.eFault;              // 非法状态拦截
    uFault := 16#0002_0317;                       // 故障级：相 ID 越界
END_CASE

(* === 段 6 · 输出映射 === *)
bError := (uFault <> 16#0000);                    // 故障标志仅由故障级码置位（R45 配对）
IF bError THEN
    uErrorId := uFault;                           // 故障级优先上报
ELSE
    uErrorId := uInfo;                            // 否则上报信息级码
END_IF
eStateOut := _eState;                             // 输出枚举段尾单点映射（N2 规则）
END_FUNCTION_BLOCK

(* ---- FB_DL_ProfinetAlarmDiag.st ---- *)
(*
    FB_DL_ProfinetAlarmDiag —— PROFINET 通道诊断聚合
    ------------------------------------------------------------------
    分类      : DL_Device / Diagnostics
    前缀      : FB_DL_
    版本      : 1.0.0
    溯源      : PROFINET 公开规范的 ChannelErrorType 枚举值（只借公开解码表，
                不解析原始诊断记录字节、不使用任何厂商诊断对象或系统库）；
                聚合结构、首出律、八类分桶、错误分级与码位 100% 自有；
                E_DL_Ne107Status 属主为 I_DL_DeviceHealth，本件只引用不重声明（R70）；
                clean-room 重写，未复制任何闭源厂商源码
    平台      : 纯 IEC 61131-3，CODESYS V3.5+ / TwinCAT 3 / InoProShop 通用
    作者      : 道莅代码库 · PLC编程专家（R19）
    ------------------------------------------------------------------
    功能说明  : 把上游已读出的通道诊断项（通道号 / 通道属性 / ChannelErrorType /
                ExtChannelErrorType / ExtChannelAddValue）分类成八类工程语义，输出故障掩码、
                首出通道、分类计数与 NE107 健康出口。本件只做语义聚合，不做字节解析。
                核心防御：① 条目数超 16 钳位处理并置故障级 0333（不越界读）；
                ② 通道号超 32767 该项跳过并计入组态错桶；
                ③ 未识别的 ChannelErrorType（含厂商自定义域）归「其他」桶并置信息码——
                   协议允许厂商自定义，未识别不等于故障；
                ④ 16#001F 语义冲突显式化：一处公开源记为临时故障，另一处记作要求维护，
                   本库按「维护类」保守侧处理并在头注释并列两种语义（不二选一硬编码）；
                ⑤ ≥ 16#8000 的系统级码（总线/同步类）不占通道掩码，单列 bSystemLevel，
                   因为运维处理路径与通道问题完全不同；
                ⑥ CASE 分类含 ELSE 兜底走「其他」桶；uEntryCount = 0 时输出全空且 eOk。
                职责边界：单通道健康判定归设备件，多源健康仲裁归 FB_DL_DeviceHealthArbiter。
    解码表    : 16#0001 短路 / 16#0002 欠压 / 16#0003 过压 / 16#0004 过载 / 16#0005 过温 /
                16#0006 断线 / 16#0007 超上限 / 16#0008 欠下限 / 16#0009 通用错误 /
                16#000F 参数缺失 / 16#0010 参数故障 / 16#001E 要求维护 / 16#001F 维护要求
                （另一公开源记为 Temporary_fault）/ >= 16#8000 系统级
    错误码    : 16#0003_016C 未识别的 ChannelErrorType（厂商自定义域），已归「其他」桶——信息级，正常防御
                16#0003_016D 预留禁用（信息级，不得挪用）
                16#0003_0333 诊断条目数超上限（> 16）——故障级，已钳位处理
                16#0003_0334 通道号越界（> 32767）——故障级，该项已跳过并计入组态错桶
                16#0003_0335 预留禁用（故障级，不得挪用）
    码位总账  : 16#0003_016C 用 / 16#0003_016D 预留 ｜ 16#0003_0333 用 / 16#0003_0334 用 / 16#0003_0335 预留
    状态机    : R6 标注 N/A —— 本组件为纯函数无顺序状态机，无 CASE 可写，非法状态不可能出现
                （分类 CASE 是协议枚举映射表，不是顺序状态机，且含 ELSE 兜底）
    采样约定  : 本件无定时器、无沿检测、无状态驻留；诊断项每拍全量重算，结论与任务周期无关。
    修订记录  : 2026-11-16 v1.0.0 首次入库（R19）
*)
FUNCTION_BLOCK FB_DL_ProfinetAlarmDiag
VAR_INPUT
    auChannelNo        : ARRAY[0..15] OF UINT;   // 通道号 [通道]，协议域 0~32767，0 表示子模块级 / channel number [channel], protocol range 0~32767, zero means submodule
    auChannelProp      : ARRAY[0..15] OF WORD;   // 通道属性（协议位域），本件原样透传不解释 [位域] / channel properties, passed through without interpretation [bitfield]
    auErrType          : ARRAY[0..15] OF WORD;   // ChannelErrorType（公开枚举，见头注释解码表）[枚举] / channel error type, see the decode table [enum]
    auExtErrType       : ARRAY[0..15] OF WORD;   // ExtChannelErrorType（厂商扩展），只透传不解释 [枚举] / extended error type, passed through only [enum]
    audAddValue        : ARRAY[0..15] OF UDINT;  // ExtChannelAddValue（附加上下文值）[无量纲] / additional context value [dimensionless]
    uEntryCount        : UINT := 0;              // 有效诊断项数 [项]，范围 0~16 / number of valid diagnostic entries [entry], range 0~16
END_VAR
VAR_OUTPUT
    uChannelMask       : WORD;                   // 有诊断的项位图，bit N = 项 N [位图] / bitmap of diagnostic entries, bit N is entry N [bitmap]
    uFirstChannel      : UINT;                   // 首出通道号（同拍取通道号最小）[通道] / first-out channel number, the lowest channel wins [channel]
    uFirstErrType      : WORD;                   // 首出项的 ChannelErrorType 原值（HMI 可查表）[枚举] / raw error type of the first-out entry [enum]
    auClassCount       : ARRAY[0..7] OF UINT;    // 八类计数 [次]，索引 0 短路 ~ 7 维护类 / eight class counters [times], 0 short circuit to 7 maintenance
    bMaintenanceOnly   : BOOL;                   // 只有维护类条目（可继续生产需保养）/ maintenance entries only, production may continue
    bSystemLevel       : BOOL;                   // 存在系统级码（>= 16#8000，总线/同步类）/ a system level code exists, bus or synchronisation class
    eHealth            : E_DL_Ne107Status;       // NE107 健康出口（引用唯一属主枚举）/ NE107 health output, referencing the owner enumeration
    eErr               : UDINT;                  // 错误码，0=正常 / error id, 0=ok
    bError             : BOOL;                   // 故障标志，eErr 为故障级时 TRUE / error flag, TRUE on fault-level eErr
    bValid             : BOOL;                   // 结论是否可用 / conclusion valid flag
END_VAR
VAR
    uIdx               : UINT;                   // 条目扫描游标 [项]，范围 0~15 / entry scan cursor [entry], range 0~15
    uCountEff          : UINT;                   // 钳位后的有效条目数 [项] / clamped effective entry count [entry]
    uClass             : UINT;                   // 本项的类别桶号 [桶]，范围 0~7 / class bucket index of this entry [bucket], range 0~7
    uBestCh            : UINT;                   // 首出通道号候选 [通道] / first-out channel candidate [channel]
    wBestErr           : WORD;                   // 首出错误类型候选 [枚举] / first-out error type candidate [enum]
    bAnyEntry          : BOOL;                   // 存在有效（占通道掩码的）条目 / at least one entry occupies the channel mask
    bUnknownType       : BOOL;                   // 本拍出现未识别的错误类型 / an unrecognised error type appeared in this cycle
    bChOutOfRange      : BOOL;                   // 本拍出现越界通道号 / an out-of-range channel number appeared in this cycle
    bFaultClass        : BOOL;                   // 存在故障类（短路~欠下限）/ a fault class entry exists
    bConfigClass       : BOOL;                   // 存在组态错类条目 / a configuration class entry exists
    bMaintainClass     : BOOL;                   // 存在维护类条目 / a maintenance class entry exists
    nChNo              : UINT;                   // 当前项的通道号（比较用副本）[通道] / channel number copy of the current entry [channel]
END_VAR
VAR CONSTANT
    DL_PN_E_SHORT       : WORD := 16#0001;       // 短路 [枚举] / short circuit [enum]
    DL_PN_E_UNDERV      : WORD := 16#0002;       // 欠压 [枚举] / undervoltage [enum]
    DL_PN_E_OVERV       : WORD := 16#0003;       // 过压 [枚举] / overvoltage [enum]
    DL_PN_E_OVERLOAD    : WORD := 16#0004;       // 过载 [枚举] / overload [enum]
    DL_PN_E_OVERTEMP    : WORD := 16#0005;       // 过温 [枚举] / overtemperature [enum]
    DL_PN_E_WIREBREAK   : WORD := 16#0006;       // 断线 [枚举] / wire break [enum]
    DL_PN_E_UPPER       : WORD := 16#0007;       // 超上限 [枚举] / upper limit exceeded [enum]
    DL_PN_E_LOWER       : WORD := 16#0008;       // 欠下限 [枚举] / lower limit violated [enum]
    DL_PN_E_GENERIC     : WORD := 16#0009;       // 通用错误 [枚举] / generic error [enum]
    DL_PN_E_PARAM_MISS  : WORD := 16#000F;       // 参数缺失 [枚举] / parameter missing [enum]
    DL_PN_E_PARAM_FAULT : WORD := 16#0010;       // 参数故障 [枚举] / parameter fault [enum]
    DL_PN_E_MAINT_REQ   : WORD := 16#001E;       // 要求维护 [枚举] / maintenance required [enum]
    DL_PN_E_MAINT_DEM   : WORD := 16#001F;       // 维护要求（另一公开源记为临时故障，本库按维护类保守处理）[枚举] / maintenance demanded, treated conservatively as maintenance [enum]
    DL_PN_E_SYS_MIN     : WORD := 16#8000;       // 系统级码起点 [枚举] / start of the system level codes [enum]
    DL_PN_CH_MAX        : UINT := 32767;         // 通道号上限 [通道] / channel number upper bound [channel]
    DL_PN_ENTRY_MAX     : UINT := 16;            // 诊断条目上限 [项] / diagnostic entry upper bound [entry]
    DL_PN_C_SHORT       : UINT := 0;             // 类别桶 0：短路 [桶] / class bucket zero, short circuit [bucket]
    DL_PN_C_WIRE        : UINT := 1;             // 类别桶 1：断线 [桶] / class bucket one, wire break [bucket]
    DL_PN_C_LOAD        : UINT := 2;             // 类别桶 2：过载 [桶] / class bucket two, overload [bucket]
    DL_PN_C_TEMP        : UINT := 3;             // 类别桶 3：过温 [桶] / class bucket three, overtemperature [bucket]
    DL_PN_C_UPPER       : UINT := 4;             // 类别桶 4：超上限 [桶] / class bucket four, upper limit [bucket]
    DL_PN_C_LOWER       : UINT := 5;             // 类别桶 5：欠下限 [桶] / class bucket five, lower limit [bucket]
    DL_PN_C_CONFIG      : UINT := 6;             // 类别桶 6：组态错/其他 [桶] / class bucket six, configuration or other [bucket]
    DL_PN_C_MAINT       : UINT := 7;             // 类别桶 7：维护类 [桶] / class bucket seven, maintenance [bucket]
    DL_PN_CLASS_CNT     : UINT := 8;             // 类别桶总数 [桶] / number of class buckets [bucket]
    DL_PN_BIT0          : WORD := 16#0001;       // 位图最低位掩码 [位图] / least significant bitmap mask [bitmap]
    DL_PN_ZERO_W        : WORD := 16#0000;       // 位图零常量 [位图] / bitmap zero constant [bitmap]
    DL_PN_ZERO          : UINT := 0;             // 无符号零常量 [无量纲] / unsigned zero constant [dimensionless]
    DL_PN_CNT_MAX       : UINT := 65535;         // 单类计数饱和值 [次] / per class counter saturation value [times]
END_VAR

// 段 1｜输出与中间量预置（位图与八类计数每拍全量重算）/ segment 1, preset outputs and intermediates
uChannelMask := DL_PN_ZERO_W;                 // 位图清零 / clear the bitmap
uFirstChannel := DL_PN_ZERO;                  // 首出通道清零 / clear the first-out channel
uFirstErrType := DL_PN_ZERO_W;                // 首出错误类型清零 / clear the first-out error type
bMaintenanceOnly := FALSE;                    // 预置非纯维护类 / preset not maintenance only
bSystemLevel := FALSE;                        // 预置无系统级码 / preset no system level code
eHealth := eOk;                               // 预置健康（条目为 0 时即为最终结论）/ preset OK, final when no entry exists
eErr := 0;                                    // 预置无错误 / preset no error
bError := FALSE;                              // 预置无故障 / preset no fault
bValid := FALSE;                              // 预置结论不可用 / preset invalid
bAnyEntry := FALSE;                           // 预置无有效条目 / preset no valid entry
bUnknownType := FALSE;                        // 预置无未识别类型 / preset no unrecognised type
bChOutOfRange := FALSE;                       // 预置无越界通道号 / preset no out-of-range channel
bFaultClass := FALSE;                         // 预置无故障类 / preset no fault class
bConfigClass := FALSE;                        // 预置无组态错类 / preset no configuration class
bMaintainClass := FALSE;                      // 预置无维护类 / preset no maintenance class
uBestCh := DL_PN_CH_MAX;                      // 首出候选初值取通道号上限（最大值哨兵）/ the candidate starts at the channel upper bound as a maximum sentinel
wBestErr := DL_PN_ZERO_W;                     // 首出错误类型初值 / initial error type of the first-out candidate
FOR uIdx := 0 TO DL_PN_CLASS_CNT - 1 DO
    auClassCount[uIdx] := DL_PN_ZERO;         // 八个类别桶逐桶清零 / clear each of the eight class buckets
END_FOR

// 段 2｜条目数闸：超上限钳位处理并置故障级（绝不越界读）/ segment 2, entry count gate
uCountEff := uEntryCount;                     // 取入参副本 / copy the input
IF uEntryCount > DL_PN_ENTRY_MAX THEN
    uCountEff := DL_PN_ENTRY_MAX;             // 钳位到 16 / clamp to sixteen
    eErr := 16#0003_0333;                     // 条目数超上限故障码 / entry count over the limit fault id
    bError := TRUE;                           // 置故障标志 / raise the error flag
END_IF

// 段 3｜零条目：协议合法（诊断记录长度 0 表示无故障）/ segment 3, zero entries is a legal protocol state
IF uCountEff = DL_PN_ZERO THEN
    eHealth := eOk;                           // 健康出口正常 / health output OK
    bValid := TRUE;                           // 结论可用 / conclusion valid
    RETURN;                                   // 无需聚合 / nothing to aggregate
END_IF

// 段 4｜逐项分类（含 ELSE 兜底走「其他」桶）/ segment 4, per entry classification
FOR uIdx := 0 TO uCountEff - 1 DO
    nChNo := auChannelNo[uIdx];               // 取本项通道号 [通道] / channel number of this entry [channel]
    IF nChNo > DL_PN_CH_MAX THEN
        bChOutOfRange := TRUE;                // 记录通道号越界 / remember the out-of-range channel
        auClassCount[DL_PN_C_CONFIG] := auClassCount[DL_PN_C_CONFIG] + 1; // 计入组态错桶 / count it in the configuration bucket
    ELSIF auErrType[uIdx] >= DL_PN_E_SYS_MIN THEN
        bSystemLevel := TRUE;                 // 系统级码单列，不占通道掩码 / system level codes are listed apart and never occupy the channel mask
    ELSE
        // 段 5｜语义分类：按公开解码表落八类桶 / segment 5, semantic classification by the public decode table
        CASE auErrType[uIdx] OF
            DL_PN_E_SHORT:
                uClass := DL_PN_C_SHORT;      // 短路 / short circuit
                bFaultClass := TRUE;          // 故障类 / fault class
            DL_PN_E_OVERV:
                uClass := DL_PN_C_UPPER;      // 过压按超上限处理 / overvoltage falls into the upper limit class
                bFaultClass := TRUE;          // 故障类 / fault class
            DL_PN_E_UNDERV:
                uClass := DL_PN_C_LOWER;      // 欠压按欠下限处理 / undervoltage falls into the lower limit class
                bFaultClass := TRUE;          // 故障类 / fault class
            DL_PN_E_WIREBREAK:
                uClass := DL_PN_C_WIRE;       // 断线 / wire break
                bFaultClass := TRUE;          // 故障类 / fault class
            DL_PN_E_OVERLOAD:
                uClass := DL_PN_C_LOAD;       // 过载 / overload
                bFaultClass := TRUE;          // 故障类 / fault class
            DL_PN_E_OVERTEMP:
                uClass := DL_PN_C_TEMP;       // 过温 / overtemperature
                bFaultClass := TRUE;          // 故障类 / fault class
            DL_PN_E_UPPER:
                uClass := DL_PN_C_UPPER;      // 超上限 / upper limit exceeded
                bFaultClass := TRUE;          // 故障类 / fault class
            DL_PN_E_LOWER:
                uClass := DL_PN_C_LOWER;      // 欠下限 / lower limit violated
                bFaultClass := TRUE;          // 故障类 / fault class
            DL_PN_E_GENERIC:
                uClass := DL_PN_C_CONFIG;     // 通用错误归其他/组态错桶 / a generic error falls into the other or configuration bucket
                bConfigClass := TRUE;         // 组态错类 / configuration class
            DL_PN_E_PARAM_MISS, DL_PN_E_PARAM_FAULT:
                uClass := DL_PN_C_CONFIG;     // 参数类一律组态错 / parameter issues are a configuration problem
                bConfigClass := TRUE;         // 组态错类 / configuration class
            DL_PN_E_MAINT_REQ, DL_PN_E_MAINT_DEM:
                uClass := DL_PN_C_MAINT;      // 维护类（16#001F 的语义冲突按保守侧归维护）/ maintenance class, the conflicting 16#001F is kept on the conservative side
                bMaintainClass := TRUE;       // 维护类 / maintenance class
        ELSE
            uClass := DL_PN_C_CONFIG;         // 未识别值归其他桶（ELSE 兜底）/ unrecognised values fall into the other bucket
            bConfigClass := TRUE;             // 组态错类 / configuration class
            bUnknownType := TRUE;             // 记录未识别类型 / remember the unrecognised type
        END_CASE

        // 段 6｜占掩码、累加计数、更新首出候选 / segment 6, occupy the mask, count and update the first-out candidate
        uChannelMask := uChannelMask OR SHL(DL_PN_BIT0, uIdx); // 置项位图，uIdx ≤ 15 移位安全 / set the entry bit, the shift never exceeds 15
        bAnyEntry := TRUE;                    // 标记存在有效条目 / flag a valid entry
        IF auClassCount[uClass] < DL_PN_CNT_MAX THEN
            auClassCount[uClass] := auClassCount[uClass] + 1; // 饱和累加，绝不回绕 / saturating increment, never wraps
        END_IF
        IF nChNo < uBestCh THEN
            uBestCh := nChNo;                 // 首出取通道号最小 / the lowest channel number wins the first-out
            wBestErr := auErrType[uIdx];      // 同步首出错误类型 / keep the matching error type
        END_IF
    END_IF
END_FOR

// 段 7｜首出发布（无有效条目则保留 0 与空类型）/ segment 7, publish the first-out
IF bAnyEntry THEN
    uFirstChannel := uBestCh;                 // 首出通道号 / first-out channel number
    uFirstErrType := wBestErr;                // 首出错误类型原值 / raw error type of the first-out entry
END_IF

// 段 8｜健康出口优先级：故障类 > 组态错 > 维护类 > 系统级 > 正常 / segment 8, health output priority
IF bFaultClass THEN
    eHealth := eFailure;                      // 短路/断线/过载/过温/越限：信号不可信 / a channel fault makes the signal untrustworthy
ELSIF bConfigClass THEN
    eHealth := eOutOfSpec;                    // 组态错：测量可能有效但不可依赖 / a configuration fault means the measurement cannot be relied upon
ELSIF bMaintainClass THEN
    eHealth := eMaintenanceReq;               // 维护类：仍有效但已劣化 / maintenance means still valid but degraded
ELSIF bSystemLevel THEN
    eHealth := eOutOfSpec;                    // 系统级：总线/同步问题，另行处理 / a system level issue is handled on a different path
ELSE
    eHealth := eOk;                           // 无任何诊断：正常 / no diagnostics, OK
END_IF

// 段 9｜纯维护类判定（可继续生产，需安排保养）/ segment 9, maintenance only evaluation
bMaintenanceOnly := bMaintainClass AND (NOT bFaultClass) AND (NOT bConfigClass); // 只有维护类条目 / maintenance entries only

// 段 10｜信息级与故障级码汇总（故障级优先，绝不互相覆盖）/ segment 10, code summary
IF bUnknownType AND (NOT bError) THEN
    eErr := 16#0003_016C;                     // 信息级：未识别类型已归其他桶 / info level, unrecognised types were bucketed as other
END_IF
IF bChOutOfRange THEN
    eErr := 16#0003_0334;                     // 通道号越界故障码 / channel number out of range fault id
    bError := TRUE;                           // 置故障标志 / raise the error flag
END_IF

// 段 11｜结论可用性（故障态仍输出分类结果供 HMI 诊断，但标记不可用于联锁）/ segment 11, conclusion validity
bValid := TRUE;                               // 分类结论本身可信（故障级只表输入越界）/ the classification itself is trustworthy, faults only mark input overruns
END_FUNCTION_BLOCK

(* ---- FB_DL_ProofTestSeq.st ---- *)
(*
  ==================================================================
  组件名 Component  : FB_DL_ProofTestSeq
  分类   Category   : DL_Device
  复杂度 Complexity  : cx4
  版本   Version    : 1.0.0
  功能   Purpose    : 联锁功能证明试验顺控。按 tTestPeriod 周期发起激励-反馈
                      回路验证：激励输出后 tFeedbackTo 内收到反馈沿进评估段，
                      保持激励 tTestDur 后按反馈在位判通过；试验失败挂
                      NE107 eCheckFunction / eMaintenanceReq 健康语言。
  来源   Source     : t2-isa-ne107（借鉴 ISA-18.2 / NE107 证明试验与健康语言
                      纪律，clean-room 自研实现，未复制任何文档代码行）
  溯源   Origin     : IEC 61131-3 标准语义的道莅防御性实现；证明试验周期激励
                      为公开功能安全维护语义。
  平台   Platform   : 纯 IEC 61131-3（Standard.library: TON / R_TRIG，无私有库）
  分工声明 Split     : 与 FB_DL_PassboxInterlockSeq（工艺顺控）分工——本件是
                      联锁回路自证试验顺控，不驱动工艺介质、不参与生产联锁。
  作者   Author     : 道莅代码库 · PLC 编程专家（R57）
  ------------------------------------------------------------------
  边界 Boundary     :
                      一 组态配比约束（R100）：tTestPeriod > tTestDur 且
                         tFeedbackTo < tTestDur，越域判故障级；
                      二 试验中真实故障（bDeviceFault）与试验失败（eTestFail）
                         分段独立成因（R190 归因唯一），真实故障优先；
                      三 试验请求仅在设备空闲相（bDevIdle）受理，运行相拒
                         并置信息级 bReqRejected 单拍；
                      四 锁存解除路径 = bReset 上升沿（唯一路径，R188）；
                      五 无全局变量、无外部变量声明、无物理地址寻址。
  修订记录 Revision  :
    2026-11-21  v1.0.0  R57 首版（批 4 · 序号 18）
  ==================================================================
*)

TYPE E_DL_PtsPhase :
(
    eIdle   := 0,  // 空闲：周期窗计时 / idle, the period window counting
    eExcite := 10, // 激励：等反馈沿 / exciting, waiting for the feedback edge
    eEval   := 20, // 评估：保持激励到持续窗满 / evaluating, the drive held until the duration expiry
    eFault  := 90  // 故障：成因锁存 / fault, the cause latched
);
END_TYPE

TYPE E_DL_PtsFault :
(
    eNone        := 0, // 无成因 / no cause
    eCfgBad      := 1, // 组态非法：三窗配比越域（故障级，与 bError 配对）/ an illegal config
    eDeviceFault := 2, // 试验中真实设备故障（故障级，与 bError 配对）/ a real device fault during the test
    eTestFail    := 3, // 试验失败：反馈超时或评估失在（故障级，与 bError 配对）/ a test failure
    ePhaseBad    := 4  // 非法相位兜底（故障级，与 bError 配对）/ an illegal phase fallback
);
END_TYPE

TYPE E_DL_PtsHealth :
(
    eGood           := 0, // NE107 正常（最近试验通过）/ the NE107 good state, the latest test passed
    eCheckFunction  := 1, // NE107 功能受影响（试验失败待复测）/ the NE107 check function state
    eMaintenanceReq := 2  // NE107 维护要求（试验失败或真实故障）/ the NE107 maintenance state
);
END_TYPE

FUNCTION_BLOCK FB_DL_ProofTestSeq
VAR_INPUT
    bEnable      : BOOL := TRUE;   // 使能，失能即停试验回空闲 [-] / enable, disabling stops the test to idle
    bReset       : BOOL := FALSE;  // 复位上升沿清锁存 [-] / reset rising edge clears the latch
    bTestReq     : BOOL := FALSE;  // 试验请求电平（仅在空闲相受理）[-] / the test request level, accepted only in idle
    bDevIdle     : BOOL := TRUE;   // 设备空闲相指示 [-] / the device idle indicator
    bDeviceFault : BOOL := FALSE;  // 设备真实故障电平 [-] / the real device fault level
    bFeedback    : BOOL := FALSE;  // 联锁反馈（激励后应动作）[-] / the interlock feedback, expected active under the drive
    tTestPeriod  : TIME := T#3600S; // 试验周期窗 [毫秒]，域 大于 tTestDur / the test period window, above the duration
    tTestDur     : TIME := T#10S;   // 试验持续窗 [毫秒]，域 大于 tFeedbackTo / the test duration window, above the feedback timeout
    tFeedbackTo  : TIME := T#5S;    // 反馈超时窗 [毫秒] / the feedback timeout window [millisecond]
END_VAR
VAR_OUTPUT
    bTestDrive   : BOOL := FALSE; // 激励输出（试验中为真）[-] / the test drive outlet
    bTestActive  : BOOL := FALSE; // 试验进行中电平 [-] / the test active level
    bTestOk      : BOOL := FALSE; // 试验通过单拍脉冲 [-] / the test pass one-scan pulse
    bReqRejected : BOOL := FALSE; // 请求被拒信息级单拍（非空闲相受理）[-] / the request rejected informational pulse
    eHealth      : E_DL_PtsHealth := E_DL_PtsHealth.eGood; // NE107 健康语言出口 [枚举] / the health outlet [enum]
    ePhase       : E_DL_PtsPhase := E_DL_PtsPhase.eIdle; // 相位出口 [枚举] / the phase outlet [enum]
    eFault       : E_DL_PtsFault := E_DL_PtsFault.eNone; // 成因出口，锁存回放 [枚举] / the cause outlet replayed
    bError       : BOOL := FALSE; // 故障锁存标志 [-] / the fault latch flag
END_VAR
VAR
    rtReset  : R_TRIG; // 复位沿检测，段 0 无条件刷新 / the reset edge
    rtReq    : R_TRIG; // 试验请求沿检测，段 0 无条件刷新 / the request edge
    rtFb     : R_TRIG; // 反馈沿检测，段 0 无条件刷新 / the feedback edge
    rtOk     : R_TRIG; // 通过电平沿检测，段 0 无条件刷新 / the pass level edge
    tonPeriod: TON;    // 试验周期窗（自复位 R188），段 0 无条件刷新 / the period window, self resetting
    tonFbTo  : TON;    // 反馈超时窗，段 0 无条件刷新 / the feedback timeout
    tonDur   : TON;    // 试验持续窗，段 0 无条件刷新 / the duration window
    _ePhase  : E_DL_PtsPhase := E_DL_PtsPhase.eIdle; // 内部相位，CASE 唯一写入目标 / the internal phase
    _eFaulC  : E_DL_PtsFault := E_DL_PtsFault.eNone; // 故障级成因，锁存至复位沿 / the fault cause, latched
    _bFault  : BOOL := FALSE; // 故障锁存位 [-] / the fault latch bit
    _bInit   : BOOL := FALSE; // 首扫初始化完成标志（R310）/ the first scan flag
    _bCfgOk  : BOOL := FALSE; // 组态域内 [-] / the config inside the domain
    _bPassed : BOOL := FALSE; // 最近试验通过保持位（复位沿清，R243 最近量）[-] / the latest pass holder, cleared by reset
END_VAR

// 段 0｜定时器与沿检测无条件周期刷新（禁入分支）/ segment 0, the unconditional refresh
rtReset(CLK := bReset); // 复位沿 / the reset edge
rtReq(CLK := bTestReq); // 请求沿 / the request edge
rtFb(CLK := bFeedback); // 反馈沿 / the feedback edge
rtOk(CLK := _bPassed); // 通过电平沿 / the pass level edge
tonPeriod(IN := bEnable AND (_ePhase = E_DL_PtsPhase.eIdle) AND (NOT tonPeriod.Q), PT := tTestPeriod); // 周期窗自复位循环（R188）/ the self resetting period loop
tonFbTo(IN := (_ePhase = E_DL_PtsPhase.eExcite) AND (NOT _bFault), PT := tFeedbackTo); // 反馈超时窗，IN 串激励相闸 / the feedback timeout gated by the excite phase
tonDur(IN := (_ePhase = E_DL_PtsPhase.eEval) AND (NOT _bFault), PT := tTestDur); // 持续窗，IN 串评估相闸 / the duration gated by the eval phase

// 段 1｜首扫初始化（R310）/ segment 1, the first scan
IF NOT _bInit THEN // 首扫一拍 / the first scan
    _bInit := TRUE; // 置首扫标志 / raise the flag
END_IF

// 段 2｜复位沿作用域：清锁存 / 清最近通过量 / 迁空闲（三项逐项声明）/ segment 2, the reset edge scope
IF rtReset.Q THEN // 复位沿 / the reset edge
    _bFault  := FALSE; // 作用域一：清故障锁存 / scope one, clear the fault latch
    _eFaulC  := E_DL_PtsFault.eNone; // 作用域一：清成因 / scope one, clear the cause
    _bPassed := FALSE; // 作用域二：清最近通过保持量（R243）/ scope two, clear the latest pass holder
    _ePhase  := E_DL_PtsPhase.eIdle; // 作用域三：迁空闲相 / scope three, back to idle
END_IF

// 段 3｜组态域闸：三窗配比（R100，边界一）/ segment 3, the config gate, the window pairing
_bCfgOk := (tTestPeriod > tTestDur) AND (tTestDur > tFeedbackTo) AND (tFeedbackTo > T#0S); // 周期 > 持续 > 反馈超时配比 / the period above duration above timeout pairing
IF NOT _bCfgOk THEN // 配比越域 / a pairing violation
    IF NOT _bFault THEN // 未锁存才迁移 / migrate only while unlatched
        _bFault := TRUE; // 置故障锁存 / raise the fault latch
        _eFaulC := E_DL_PtsFault.eCfgBad; // 故障级成因（R45 配对 bError）/ the fault cause
        _ePhase := E_DL_PtsPhase.eFault; // 迁故障相 / migrate to fault
    END_IF
END_IF

// 段 4｜相位机：ENUM + CASE，含 ELSE 非法相位兜底（R128）/ segment 4, the phase machine
CASE _ePhase OF

E_DL_PtsPhase.eIdle: // 空闲相：请求受理与周期触发 / the idle phase, the request acceptance and the period trigger
    IF NOT bEnable THEN // 失能 / disabled
        _ePhase := E_DL_PtsPhase.eIdle; // 停摆驻留 / dwell
    ELSIF rtReq.Q AND (NOT bDevIdle) THEN // 非空闲相受理请求（边界三）/ a request while not idle
        bReqRejected := TRUE; // 信息级拒绝单拍 / the informational reject pulse
    ELSIF (tonPeriod.Q OR rtReq.Q) AND bDevIdle AND (NOT _bFault) THEN // 周期到或请求沿且空闲 / the period expiry or an accepted request
        _ePhase := E_DL_PtsPhase.eExcite; // 迁激励相 / migrate to excite
    END_IF

E_DL_PtsPhase.eExcite: // 激励相：等反馈沿 / the excite phase, waiting for the feedback edge
    IF NOT bEnable THEN // 失能 / disabled
        _ePhase := E_DL_PtsPhase.eIdle; // 回空闲相 / back to idle
    ELSIF bDeviceFault THEN // 真实故障优先（边界二）/ the real fault first
        _bFault := TRUE; // 置故障锁存 / raise the fault latch
        _eFaulC := E_DL_PtsFault.eDeviceFault; // 故障级成因（R45 配对 bError）/ the fault cause
        _ePhase := E_DL_PtsPhase.eFault; // 迁故障相 / migrate to fault
    ELSIF rtFb.Q THEN // 反馈沿到达 / a feedback edge arrived
        _ePhase := E_DL_PtsPhase.eEval; // 迁评估相 / migrate to eval
    ELSIF tonFbTo.Q THEN // 反馈超时 / the feedback timed out
        _bFault := TRUE; // 置故障锁存 / raise the fault latch
        _eFaulC := E_DL_PtsFault.eTestFail; // 故障级成因（R45 配对 bError）/ the fault cause
        _ePhase := E_DL_PtsPhase.eFault; // 迁故障相 / migrate to fault
    END_IF

E_DL_PtsPhase.eEval: // 评估相：保持激励到持续窗满再判反馈在位 / the eval phase, the drive held then the verdict
    IF NOT bEnable THEN // 失能 / disabled
        _ePhase := E_DL_PtsPhase.eIdle; // 回空闲相 / back to idle
    ELSIF bDeviceFault THEN // 真实故障优先（边界二）/ the real fault first
        _bFault := TRUE; // 置故障锁存 / raise the fault latch
        _eFaulC := E_DL_PtsFault.eDeviceFault; // 故障级成因（R45 配对 bError）/ the fault cause
        _ePhase := E_DL_PtsPhase.eFault; // 迁故障相 / migrate to fault
    ELSIF tonDur.Q THEN // 持续窗满 / the duration expired
        IF bFeedback THEN // 反馈在位判通过 / the feedback held, a pass
            _bPassed := TRUE; // 置最近通过保持量 / raise the pass holder
        ELSE // 反馈脱落判失败 / the feedback dropped, a failure
            _bFault := TRUE; // 置故障锁存 / raise the fault latch
            _eFaulC := E_DL_PtsFault.eTestFail; // 故障级成因（R45 配对 bError）/ the fault cause
            _ePhase := E_DL_PtsPhase.eFault; // 迁故障相 / migrate to fault
        END_IF
        IF NOT _bFault THEN // 通过路径回空闲 / the pass path back to idle
            _ePhase := E_DL_PtsPhase.eIdle; // 回空闲相 / back to idle
        END_IF
    END_IF

E_DL_PtsPhase.eFault: // 故障相：成因锁存，等复位沿；失能也回空闲（解锁路径，R188）/ the fault phase, latched until the reset edge
    IF NOT bEnable THEN // 失能 / disabled
        _ePhase := E_DL_PtsPhase.eIdle; // 回空闲相（锁存仍保持至复位沿）/ back to idle, the latch held until reset
    END_IF

ELSE // 非法相位兜底（R128）/ the illegal phase fallback
    _bFault := TRUE; // 置故障锁存 / raise the fault latch
    _eFaulC := E_DL_PtsFault.ePhaseBad; // 故障级成因（R45 配对 bError）/ the fault cause
    _ePhase := E_DL_PtsPhase.eFault; // 迁故障相 / migrate to fault
END_CASE

// 段 5｜统一出口 / segment 5, the unified outlet
bTestDrive := (_ePhase = E_DL_PtsPhase.eExcite) OR (_ePhase = E_DL_PtsPhase.eEval); // 激励输出（激励与评估相保持）/ the drive held in excite and eval
bTestActive := bTestDrive; // 试验进行中电平 / the active level
bTestOk := rtOk.Q; // 通过单拍脉冲（沿检测已无条件刷新）/ the pass pulse
IF _bFault THEN // 故障锁存优先 / the fault latch first
    eFault := _eFaulC; // 成因锁存回放（R152）/ the cause replayed
    IF _eFaulC = E_DL_PtsFault.eTestFail THEN // 试验失败映射功能受影响（NE107）/ a test failure maps to check function
        eHealth := E_DL_PtsHealth.eCheckFunction; // 功能受影响 / the check function state
    ELSE // 其余故障映射维护要求 / the other causes to maintenance
        eHealth := E_DL_PtsHealth.eMaintenanceReq; // 维护要求 / the maintenance state
    END_IF
ELSE // 无锁存 / no latch
    eFault := E_DL_PtsFault.eNone; // 无成因 / no cause
    eHealth := E_DL_PtsHealth.eGood; // 健康态 / the good state
END_IF
ePhase := _ePhase; // 相位出口单点映射 / the phase outlet
bError := _bFault; // 故障标志与锁存位同源 / the flag shares the latch
END_FUNCTION_BLOCK
